// TIA Portal V20 program export: 0 tag tables, 0 data types, 52 data blocks, 105 code blocks (in call order from the OBs), 282 instance data blocks

DATA_BLOCK "Bypass"   // DB9
{ S7_Optimized_Access := 'TRUE' }
VERSION : 0.1
// stored: AutoNumber true, DBAccessibleFromOPCUA true, IsOnlyStoredInLoadMemory false, IsRetainMemResEnabled false, IsWriteProtectedInAS false, MemoryReserve 100
   VAR RETAIN
      Main_Panel { S7_SetPoint := 'True'} : "Safety_Bypass_MainPanel";
      Remote_Panel_1 : "Safety_Bypass_RemotePanel";
      Remote_Panel_2 { S7_SetPoint := 'True'} : "Safety_Bypass_RemotePanel";
      Remote_Panel_3 { S7_SetPoint := 'True'} : "Safety_Bypass_RemotePanel";
      Remote_Panel_4 { S7_SetPoint := 'True'} : "Safety_Bypass_RemotePanel";
      Remote_Panel_5 { S7_SetPoint := 'True'} : "Safety_Bypass_RemotePanel";
   END_VAR
BEGIN
   Main_Panel.Estop_Cabinet := FALSE;
END_DATA_BLOCK

DATA_BLOCK "Bypass_Safe"   // DB39, F_DB
{ S7_Optimized_Access := 'TRUE' }
VERSION : 0.1
// stored: AutoNumber true, DBAccessibleFromOPCUA true
   VAR
      Main_Panel : "F_Bypass_MainPanel";
      Remote_Panel_1 : "F_Bypass_RemotePanel";
      Remote_Panel_2 : "F_Bypass_RemotePanel";
      Remote_Panel_3 : "F_Bypass_RemotePanel";
      Remote_Panel_4 : "F_Bypass_RemotePanel";
      Remote_Panel_5 : "F_Bypass_RemotePanel";
   END_VAR
BEGIN
END_DATA_BLOCK

DATA_BLOCK "CNV_HMI"   // DB40
{ S7_Optimized_Access := 'TRUE' }
VERSION : 0.1
// stored: AutoNumber true, DBAccessibleFromOPCUA true, IsOnlyStoredInLoadMemory false, IsRetainMemResEnabled false, IsWriteProtectedInAS false, MemoryReserve 100
   VAR
      "Manual_Sfty_Stopper_Up(1)" : Array[1..5] of Bool;
      "Manual_Sfty_Stopper_Down(1)" : Array[1..5] of Bool;
      In_Out : Array[1..5] of Bool;
      ID : Array[1..5] of DInt;
      "Task_ID(1)" : Array[1..5] of UInt;
      Manual_Bwd : Array[1..5] of Bool;
      "Reset(1)" : Array[1..5] of Bool;
      "Pallet_Type(1)" : Array[1..5] of UInt;
      Manual_Fwd : Array[1..5] of Bool;
      Enable : Array[1..5] of Bool;
      "Pallet_Align_Right(1)" : Array[1..5] of Bool;
      "Enable(1)" : Array[1..5] of Bool;
      Pallet_Type : Array[1..5] of UInt;
      Pallet_Allignment : Array[1..5] of Bool;
      "Transfer_To_ID(1)" : Array[1..5] of DInt;
      Pallet_Align_Right : Array[1..5] of Bool;
      "Manual_Bwd(1)" : Array[1..5] of Bool;
      "Pallet_Align_Left(1)" : Array[1..5] of Bool;
      Reset : Array[1..5] of Bool;
      Stop : Array[1..5] of Bool;
      Pallet_Align_Center : Array[1..5] of Bool;
      "Stop(1)" : Array[1..5] of Bool;
      "Start_Transfer(1)" : Array[1..5] of Bool;
      Pallet_Align_Left : Array[1..5] of Bool;
      Start_Transfer : Array[1..5] of Bool;
      "ID(1)" : Array[1..5] of DInt;
      "Transfer_From_ID(1)" : Array[1..5] of DInt;
      "Manual_Fwd(1)" : Array[1..5] of Bool;
      Mode_Change : Array[1..5] of UInt;
      Transfer_To_ID : Array[1..5] of DInt;
      "Mode_Change(1)" : Array[1..5] of UInt;
      Transfer_From_ID : Array[1..5] of DInt;
      UpDown : Array[1..5] of UInt;
      Same_Cnv : Array[1..5] of Bool;
      CNV2_Selected : Array[1..5] of UInt;
      "Pallet_Allignment(1)" : Array[1..5] of Bool;
      "Occupied(1)" : Array[1..5] of Bool;
      Mode : Array[1..5] of UInt;
      "Running(1)" : Array[1..5] of Bool;
      "Enabled(1)" : Array[1..5] of Bool;
      Motor_Speed_Actual : Array[1..5] of UInt;
      Running : Array[1..5] of Bool;
      "SM_State(1)" : Array[1..5] of UInt;
      "Warning(1)" : Array[1..5] of UInt;
      Stopped : Array[1..5] of Bool;
      Enabled : Array[1..5] of Bool;
      Error : Array[1..5] of Bool;
      "Motor_Speed_Requested(1)" : Array[1..5] of UInt;
      Current_Task_ID : Array[1..5] of UInt;
      "Mode(1)" : Array[1..5] of UInt;
      "Current_Task_Type(1)" : Array[1..5] of UInt;
      Warning : Array[1..5] of UInt;
      "Current_Task_ID(1)" : Array[1..5] of UInt;
      Current_Task_Type : Array[1..5] of UInt;
      "Stopped(1)" : Array[1..5] of Bool;
      Motor_Direction : Array[1..5] of UInt;
      SM_State : Array[1..5] of UInt;
      "Ready_For_Task(1)" : Array[1..5] of Bool;
      Ready_For_Task : Array[1..5] of Bool;
      Occupied : Array[1..5] of Bool;
      "Error(1)" : Array[1..5] of Bool;
      Shuttle_in_place : Array[1..5] of Bool;
      Motor_Speed_Requested : Array[1..5] of UInt;
      "Motor_Direction(1)" : Array[1..5] of UInt;
      "Motor_Speed_Actual(1)" : Array[1..5] of UInt;
      "Shuttle_in_place(1)" : Array[1..5] of Bool;
      Motor_Ready : Array[1..5] of Bool;
      "Motor_Current_Actual(1)" : Array[1..5] of Real;
      Motor_Status : Array[1..5] of UInt;
      "Motor_Status(1)" : Array[1..5] of UInt;
      Motor_Current_Actual : Array[1..5] of Real;
      "Motor_Ready(1)" : Array[1..5] of Bool;
      Task_ID : Array[1..5] of UInt;
      Level_Selected : Array[1..5] of UInt;
      "UpDown(1)" : Array[1..5] of UInt;
      Motor_Actual_Torque : Array[1..5] of Real;
      "Motor_Actual_Torque(1)" : Array[1..5] of Real;
      Safety_OK : Array[1..5] of Bool;
      Reset_Comissioning : Array[1..5] of Bool;
      Charge_Commands : Array[1..5] of Bool;
      Charge_Cnv : Array[1..5] of Bool;
      Reset_All : Array[1..5] of Bool;
      Sdetect1 : Array[1..5] of Bool;
      Sdetect2 : Array[1..5] of Bool;
      "Sdetect1(1)" : Array[1..5] of Bool;
      "Sdetect2(1)" : Array[1..5] of Bool;
      "Rpd2(1)" : Array[1..5] of Bool;
      Center : Array[1..5] of Bool;
      "Rpd1(1)" : Array[1..5] of Bool;
      "Lpd2(1)" : Array[1..5] of Bool;
      "Lpd1(1)" : Array[1..5] of Bool;
      Rpd1 : Array[1..5] of Bool;
      Lpd1 : Array[1..5] of Bool;
      Rpd2 : Array[1..5] of Bool;
      "Right(1)" : Array[1..5] of Bool;
      Right : Array[1..5] of Bool;
      Left : Array[1..5] of Bool;
      "Left(1)" : Array[1..5] of Bool;
   END_VAR
BEGIN
END_DATA_BLOCK

DATA_BLOCK "Control_DB"   // DB69
{ S7_Optimized_Access := 'TRUE' }
VERSION : 0.1
// stored: AutoNumber true, DBAccessibleFromOPCUA true, IsOnlyStoredInLoadMemory false, IsRetainMemResEnabled false, IsWriteProtectedInAS false, MemoryReserve 100
   VAR
      ECnv_Sys { S7_SetPoint := 'True'} : Array[1..5] of "ECnv_Control";
      LCnv_Sys { S7_SetPoint := 'True'} : Array[1..5] of "Cnv_VTD_Control";
      VTD_Sys { S7_SetPoint := 'True'} : Array[1..5] of "VTD_Control";
      WCS_OPC_Control { S7_SetPoint := 'True'} : Array[1..5] of "WMS_OPC_UA";
      Shuttles_Position : Array[1..23] of Struct
         x : DInt;
         y : DInt;
         Charging : Bool;
      END_STRUCT;
      VTDBarcode_Station : Array[1..5] of "Barcode_Station_UDT";
      Pallet_ID_Received : Array[1..3] of Bool;
      Gate_Station : Array[1..12] of "Gate_Station_UDT";
   END_VAR
BEGIN
   LCnv_Sys[4].Cnv_Level[1..8].Cnv2.Safety_Stop_Cnrl.Inputs.DP_Extended := TRUE;
   LCnv_Sys[5].Cnv_Level[1..8].Cnv2.Safety_Stop_Cnrl.Inputs.DP_Extended := TRUE;
END_DATA_BLOCK

DATA_BLOCK "DB_Receive_Data_From_Logistex"   // DB900
{ S7_Optimized_Access := 'TRUE' }
VERSION : 0.1
// stored: AutoNumber false, DBAccessibleFromOPCUA true, IsOnlyStoredInLoadMemory false, IsRetainMemResEnabled false, IsWriteProtectedInAS false, MemoryReserve 100
   VAR
      J1310_Conv_Infeed : "Conv_Infeed";
      J1320_Conv_Infeed { S7_SetPoint := 'True'} : "Conv_Infeed";
      J1330_Conv_Infeed { S7_SetPoint := 'True'} : "Conv_Infeed";
      J1310_Conv_Oufeed { S7_SetPoint := 'True'} : "Conv_Outfeed";
      J1320_Conv_Oufeed { S7_SetPoint := 'True'} : "Conv_Outfeed";
      J1330_Conv_Oufeed { S7_SetPoint := 'True'} : "Conv_Outfeed";
      CNV_STATUS : Array[1..10] of Byte;
      PLC_STATUS : Struct
         Hardbit : Bool;
         "PLC_E-Stop" : Bool;
      END_STRUCT;
   END_VAR
BEGIN
END_DATA_BLOCK

DATA_BLOCK "DB_Send_Data_To_Logistex"   // DB901
{ S7_Optimized_Access := 'TRUE' }
VERSION : 0.1
// stored: AutoNumber false, DBAccessibleFromOPCUA true, IsOnlyStoredInLoadMemory false, IsRetainMemResEnabled false, IsWriteProtectedInAS false, MemoryReserve 100
   VAR
      VTD_J1310_INFEED : "VTD_Infeed";
      VTD_J1320_INFEED { S7_SetPoint := 'True'} : "VTD_Infeed";
      VTD_J1330_INFEED { S7_SetPoint := 'True'} : "VTD_Infeed";
      VTD_J1310_OUTFEED { S7_SetPoint := 'True'} : "VTD_Outfeed";
      VTD_J1320_OUTFEED { S7_SetPoint := 'True'} : "VTD_Outfeed";
      VTD_J1330_OUTFEED { S7_SetPoint := 'True'} : "VTD_Outfeed";
      VTD_STATUS : Array[1..10] of Byte;
      PLC_STATUS : Struct
         Hardbit : Bool;
         "PLC_E-Stop" : Bool;
      END_STRUCT;
      CONV_SPEED : Struct
         VTD_J1310_INF_SP : Int;
         VTD_J1310_OUF_SP : Int;
         VTD_J1320_INF_SP : Int;
         VTD_J1320_OUF_SP : Int;
         VTD_J1330_INF_SP_1 : Int;
         VTD_J1330_OUF_SP : Int;
      END_STRUCT;
   END_VAR
BEGIN
END_DATA_BLOCK

DATA_BLOCK "Force"   // DB12
{ S7_Optimized_Access := 'TRUE' }
VERSION : 0.1
// stored: AutoNumber true, DBAccessibleFromOPCUA true, IsOnlyStoredInLoadMemory false, IsRetainMemResEnabled false, IsWriteProtectedInAS false, MemoryReserve 100
   VAR
      "MAIN PANEL STACK LIGHT RED" : Bool;
      "MAIN PANEL STACK LIGHT AMBER" : Bool;
      "MAIN PANEL STACK LIGHT GREEN" : Bool;
      Remote_Panel : Array[1..5] of Struct
         "CX101_SFTY STOPPER ROTATE" : Bool;
         "CX102_SFTY STOPPER ROTATE" : Bool;
         "CX103_SFTY STOPPER ROTATE" : Bool;
         "CX104_SFTY STOPPER ROTATE" : Bool;
         "CX105_SFTY STOPPER ROTATE" : Bool;
         "CX106_SFTY STOPPER ROTATE" : Bool;
         "CX107_SFTY STOPPER ROTATE" : Bool;
         "CX108_SFTY STOPPER ROTATE" : Bool;
         "CX201_SFTY STOPPER ROTATE" : Bool;
         "CX202_SFTY STOPPER ROTATE" : Bool;
         "CX203_SFTY STOPPER ROTATE" : Bool;
         "CX204_SFTY STOPPER ROTATE" : Bool;
         "CX205_SFTY STOPPER ROTATE" : Bool;
         "CX206_SFTY STOPPER ROTATE" : Bool;
         "CX207_SFTY STOPPER ROTATE" : Bool;
         "CX208_SFTY STOPPER ROTATE" : Bool;
         "VTDx DOCKING PINS 1 RETRACT" : Bool;
         "VTDx DOCKING PINS 1 EXTEND" : Bool;
         "VTDx DOCKING PINS 2 EXTEND" : Bool;
         "VTDx DOCKING PINS 2 RETRACT" : Bool;
         "SCA X00Y STACK LIGHTS AMBER" : Bool;
         "SCA X00Y STACK LIGHTS GREEN" : Bool;
         "SCA X00Y STACK LIGHTS RED" : Bool;
         "EMERGENCY STOP RESET STATUS - ON(X)" : Bool;
      END_STRUCT;
   END_VAR
BEGIN
END_DATA_BLOCK

DATA_BLOCK "HMI_DB"   // DB21
{ S7_Optimized_Access := 'TRUE' }
VERSION : 0.1
// stored: AutoNumber true, DBAccessibleFromOPCUA true, IsOnlyStoredInLoadMemory false, IsRetainMemResEnabled false, IsWriteProtectedInAS false, MemoryReserve 100
   VAR
      Username : String := 'admin';
      Password : String := '12345';
      ScreenNo : Array[1..5] of UInt;
      ScreenNo_Main : UInt;
      System_Selected : Array[1..5] of UInt;
      Rem_Loc_Keys { ExternalAccessible := 'False'; ExternalVisible := 'False'; ExternalWritable := 'False'} : Array[1..5] of "Level_Keys_UDT";
   END_VAR
BEGIN
END_DATA_BLOCK

DATA_BLOCK "HMI_OrderTable"   // DB110
{ S7_Optimized_Access := 'TRUE' }
VERSION : 0.1
// stored: AutoNumber true, DBAccessibleFromOPCUA true, IsOnlyStoredInLoadMemory false, IsRetainMemResEnabled false, IsWriteProtectedInAS false, MemoryReserve 100
   VAR
      OrderTable : Array[0..9] of "OrderTable_UDT";
      State { S7_SetPoint := 'True'} : Array[0..9] of USInt;
      Index : Array[0..9] of Int;
      ScrollUp_PB : Bool;
      ScrollDown_PB : Bool;
      PlaceOrder_PB : Bool;
      PauseOrders_PB : Bool;
      ResumeOrder_PB : Bool;
      CancelOrder_PB : Bool;
      CancelThisOrder_PB : Bool;
      StartRow : Int;
      Device : USInt;
      PlacingNewOrder : Bool;
      PopUp_ErrorWindow_Active : Bool;
      PopUp_ErrorID : UInt;
      PopUp_Index : Int;
   END_VAR
BEGIN
END_DATA_BLOCK

DATA_BLOCK "HMI_OrderTable_1"   // DB137
{ S7_Optimized_Access := 'TRUE' }
VERSION : 0.1
// stored: AutoNumber true, DBAccessibleFromOPCUA true, IsOnlyStoredInLoadMemory false, IsRetainMemResEnabled false, IsWriteProtectedInAS false, MemoryReserve 100
   VAR
      OrderTable : Array[0..9] of "OrderTable_UDT";
      State { S7_SetPoint := 'True'} : Array[0..9] of USInt;
      Index : Array[0..9] of Int;
      ScrollUp_PB : Bool;
      ScrollDown_PB : Bool;
      PlaceOrder_PB : Bool;
      PauseOrders_PB : Bool;
      ResumeOrder_PB : Bool;
      CancelOrder_PB : Bool;
      CancelThisOrder_PB : Bool;
      StartRow : Int;
      Device : USInt;
      PlacingNewOrder : Bool;
      PopUp_ErrorWindow_Active : Bool;
      PopUp_ErrorID : UInt;
      PopUp_Index : Int;
   END_VAR
BEGIN
END_DATA_BLOCK

DATA_BLOCK "OrderTable_HMI"   // DB96
{ S7_Optimized_Access := 'TRUE' }
VERSION : 0.1
// stored: AutoNumber true, DBAccessibleFromOPCUA true, IsOnlyStoredInLoadMemory false, IsRetainMemResEnabled false, IsWriteProtectedInAS false, MemoryReserve 100
   VAR
      Start : Bool;
      Pause : Bool;
      Resume : Bool;
      Stop : Bool;
      "Manual order" : Bool;
      Transfer_From_To : Byte;
      "Send VTD Order" : Bool;
      "Send CNV Order" : Bool;
      "Pallet Type" : Byte;
      "Tower 1 Pallet Alignment" : Byte;
      "Tower 2 Pallet Alignment" : Byte;
      "Extractor Pallet Alignment" : Byte;
      "From level" : Byte;
      "To level" : Byte;
      "Testing Time" : UInt;
      "Numer of cycles" : Byte;
      Tower : Byte;
      Level : Byte;
      "Time Running" : UInt;
      Actual_Cycle : Byte;
      "Start Test Visibility" : Bool;
      "Stop Test Visibility" : Bool;
      "Pause Test Visibility" : Bool;
      "Resume Visibility" : Bool;
      "Clear Table Visibility" : Bool;
      "Pallet Type Visibility" : Bool;
      "Tower 1 Visibility" : Bool;
      "Tower 2 Visibility" : Bool;
      "Extractor Visibility" : Bool;
      Auto_Settings_Visibility : Bool;
      "ToExtractor Visibility" : Bool;
      "Manual order Visibility" : Bool;
      "Tower Visibility" : Bool;
      "Level Visibility" : Bool;
      "Send VTD Order Visibility" : Bool;
      "Send CNV Order Visibility" : Bool;
   END_VAR
BEGIN
END_DATA_BLOCK

DATA_BLOCK "OrderTable_HMI_1"   // DB99
{ S7_Optimized_Access := 'TRUE' }
VERSION : 0.1
// stored: AutoNumber true, DBAccessibleFromOPCUA true, IsOnlyStoredInLoadMemory false, IsRetainMemResEnabled false, IsWriteProtectedInAS false, MemoryReserve 100
   VAR
      Start : Bool;
      Pause : Bool;
      Resume : Bool;
      Stop : Bool;
      "Manual order" : Bool;
      Transfer_From_To : Byte;
      "Send VTD Order" : Bool;
      "Send CNV Order" : Bool;
      "Pallet Type" : Byte;
      "Tower 1 Pallet Alignment" : Byte;
      "Tower 2 Pallet Alignment" : Byte;
      "Extractor Pallet Alignment" : Byte;
      "From level" : Byte;
      "To level" : Byte;
      "Testing Time" : UInt;
      "Numer of cycles" : Byte;
      Tower : Byte;
      Level : Byte;
      "Time Running" : UInt;
      Actual_Cycle : Byte;
      "Start Test Visibility" : Bool;
      "Stop Test Visibility" : Bool;
      "Pause Test Visibility" : Bool;
      "Resume Visibility" : Bool;
      "Clear Table Visibility" : Bool;
      "Pallet Type Visibility" : Bool;
      "Tower 1 Visibility" : Bool;
      "Tower 2 Visibility" : Bool;
      "Extractor Visibility" : Bool;
      Auto_Settings_Visibility : Bool;
      "ToExtractor Visibility" : Bool;
      "Manual order Visibility" : Bool;
      "Tower Visibility" : Bool;
      "Level Visibility" : Bool;
      "Send VTD Order Visibility" : Bool;
      "Send CNV Order Visibility" : Bool;
      Clear_OT : Bool;
   END_VAR
BEGIN
END_DATA_BLOCK

DATA_BLOCK "Overhang_IO_DB"   // DB439, F_DB
{ S7_Optimized_Access := 'TRUE' }
VERSION : 0.1
// stored: AutoNumber true, DBAccessibleFromOPCUA true
   VAR
      ECnv_1 : "F_ECnv_Overhang";
      ECnv_2 : "F_ECnv_Overhang";
      ECnv_3 : "F_ECnv_Overhang";
      ECnv_4 : "F_ECnv_Overhang";
      ECnv_5 : "F_ECnv_Overhang";
   END_VAR
BEGIN
END_DATA_BLOCK

DATA_BLOCK "PopUp_Screens_1"   // DB51
{ S7_Optimized_Access := 'TRUE' }
VERSION : 0.1
// stored: AutoNumber true, DBAccessibleFromOPCUA true, IsOnlyStoredInLoadMemory false, IsRetainMemResEnabled false, IsWriteProtectedInAS false, MemoryReserve 100
   VAR
      LE_Speed : Array[1..6] of DInt;
      LE_Warnings : Array[1..6] of Byte;
      LE_Status : Array[1..6] of Bool;
      LE_Quality_Value : Array[1..6] of Int;
      LE_X_Unsafe_Position : Array[1..6] of UInt;
      LE_Quality_Decoded_Codes : Array[1..6] of UInt;
      LE_Bypass : Array[1..6] of DInt;
      AE_Speed : Array[1..6] of DInt;
      AE_Status_2 : Array[1..6] of UInt;
      AE_Control_Word_2 : Array[1..6] of UInt;
      AE_Position_1 : Array[1..6] of Bool;
      AE_Position_2 : Array[1..6] of Bool;
      AE_Status_1 : Array[1..6] of Bool;
      AE_Control_Word_1 : Array[1..6] of Bool;
      BCD_Disable_Trigger_HMI : Array[1..6] of Bool;
      BCD_Enable_Trigger_HMI : Array[1..6] of Bool;
      BCD_Error_HMI : Array[1..6] of Bool;
      BCD_Start_Comm_Test_HMI : Array[1..6] of Bool;
      BCD_Test_Ok_HMI : Array[1..6] of Bool;
      BCD_Execute_Function : Array[1..6] of Bool;
      BCD_RdDone : Array[1..6] of Bool;
      BCD_ReqDone : Array[1..6] of Bool;
      BCD_ReqBusy : Array[1..6] of Bool;
   END_VAR
BEGIN
END_DATA_BLOCK

DATA_BLOCK "PopUps_DB"   // DB38
{ S7_Optimized_Access := 'TRUE' }
VERSION : 0.1
// stored: AutoNumber false, DBAccessibleFromOPCUA true, IsOnlyStoredInLoadMemory false, IsRetainMemResEnabled false, IsWriteProtectedInAS false, MemoryReserve 100
   VAR
      Buffer_Cnv_Settings_1 : "Buffer_Cnv_Settings";
      Buffer_Cnv_Settings_2 { S7_SetPoint := 'True'} : "Buffer_Cnv_Settings";
      ECnv_Settings { S7_SetPoint := 'True'} : "ECnv_Settings";
      VTD_Settings { S7_SetPoint := 'True'} : "VTD_Settings";
      Shuttle_MQTT_Settings { S7_SetPoint := 'True'} : "MQTT_Settings";
      Sick_Lector_Reseult : String;
   END_VAR
BEGIN
END_DATA_BLOCK

DATA_BLOCK "PopUps_DB_1"   // DB20
{ S7_Optimized_Access := 'TRUE' }
VERSION : 0.1
// stored: AutoNumber true, DBAccessibleFromOPCUA true, IsOnlyStoredInLoadMemory false, IsRetainMemResEnabled false, IsWriteProtectedInAS false, MemoryReserve 100
   VAR
      Buffer_Cnv_Settings_1 : Array[1..5] of "Buffer_Cnv_Settings";
      Buffer_Cnv_Settings_2 { S7_SetPoint := 'True'} : Array[1..5] of "Buffer_Cnv_Settings";
      ECnv_Settings { S7_SetPoint := 'True'} : Array[1..5] of "ECnv_Settings";
      VTD_Settings { S7_SetPoint := 'True'} : Array[1..5] of "VTD_Settings";
      Shuttle_MQTT_Settings { S7_SetPoint := 'True'} : "MQTT_Settings";
      Sick_Lector_Reseult : Array[1..5] of String;
      Save_Settings { S7_SetPoint := 'True'} : Array[1..5] of Bool;
      Absolute_Encoder : Array[1..5] of Struct
         AE_Control_Word_1 : UInt;
         AE_Control_Word_2 : UInt;
         AE_Status_1 : UInt;
         AE_Status_2 : UInt;
         AE_Position_1 : DInt;
         AE_Position_2 : DInt;
         AE_Speed : Int;
      END_STRUCT;
      Lector_Barcode : Array[1..5] of Struct
         BCD_Test_Comm : Bool;
         BCD_Disable_Trigger : Bool;
         BCD_Enable_Trigger : Bool;
         BCD_Execute_Function : Bool;
         BCD_Test_Ok : Bool;
         BCD_Error : Bool;
         BCD_RdDone : Bool;
         BCD_ReqDone : Bool;
         BCD_ReqBusy : Bool;
         Lector_Reseult : String;
      END_STRUCT;
      Linear_Encoder : Array[1..5] of Struct
         LE_X_Unsafe_Position : DInt;
         LE_Speed : Int;
         LE_Warnings : Int;
         LE_Bypass : Bool;
         LE_Status : UInt;
      END_STRUCT;
      Trend : Array[1..5] of Struct
         Motor_SetPoint : UInt;
         Motor_Actual_Current : Real;
         Motor_Actual_Speed : UInt;
      END_STRUCT;
   END_VAR
BEGIN
   Shuttle_MQTT_Settings.MQTT_Con_Params.hwId := 64;
   Shuttle_MQTT_Settings.MQTT_Con_Params.broker := '10.0.34.2';
   Shuttle_MQTT_Settings.Client_ID := WSTRING#'PLC';
   Shuttle_MQTT_Settings.Username := WSTRING#'Devin';
   Shuttle_MQTT_Settings.Password := WSTRING#'1';
   Shuttle_MQTT_Settings.Retain := TRUE;
END_DATA_BLOCK

DATA_BLOCK "SICK_AFx60_Data_DB"   // DB120
{ S7_Optimized_Access := 'TRUE' }
VERSION : 0.1
// stored: AutoNumber true, DBAccessibleFromOPCUA true, IsOnlyStoredInLoadMemory false, IsRetainMemResEnabled false, IsWriteProtectedInAS false, MemoryReserve 100
   VAR
      "Absolute Encoder 1" { S7_SetPoint := 'True'} : "ST_SICK_AFx60";
      "Absolute Encoder 2" { S7_SetPoint := 'True'} : "ST_SICK_AFx60";
      "Absolute Encoder 3" { S7_SetPoint := 'True'} : "ST_SICK_AFx60";
      "Absolute Encoder 4" { S7_SetPoint := 'True'} : "ST_SICK_AFx60";
      "Absolute Encoder 5" { S7_SetPoint := 'True'} : "ST_SICK_AFx60";
   END_VAR
BEGIN
END_DATA_BLOCK

DATA_BLOCK "SICK_Lector_DB_1"   // DB46
{ S7_Optimized_Access := 'TRUE' }
VERSION : 0.1
// stored: AutoNumber true, DBAccessibleFromOPCUA true, IsOnlyStoredInLoadMemory false, IsRetainMemResEnabled false, IsWriteProtectedInAS false, MemoryReserve 100
   VAR
      Barcode_Result : String;
      Test_OK : Bool;
      HWInputIdent : HW_IO := 554;
      HWInputLength : USInt := 32;
      HWOutputIdent : HW_IO := 555;
      HWOutputLength : USInt := 32;
      CANId : USInt := 0;
      TOut : Time := T#10S;
      Req : Bool := FALSE;
      TriggerOn : Bool := FALSE;
      TriggerOff : Bool := FALSE;
      Matchcode : Bool := FALSE;
      SavePermanent : Bool := FALSE;
      ComTest : Bool := FALSE;
      FreeCommand : Bool := FALSE;
      Data : "ST_SICK_Lector_CLV6xx";
      RdDone { S7_SetPoint := 'True'} : Bool := FALSE;
      ReqDone : Bool := FALSE;
      ReqBusy : Bool := FALSE;
      Error : Bool := TRUE;
      Errorcode : DWord := 16#0000_0015;
   END_VAR
BEGIN
   Data.Matchcode.sName := '';
   Data.Matchcode.nCodeType := ' ';
   Data.Matchcode.iMinMaxLength := 0;
   Data.Matchcode.sContent := '';
   Data.FreeCommand.sCommand := '';
   Data.FreeCommand.sResult := '';
   Data.ReadingResult.iCounter := 0;
   Data.ReadingResult.iLength := 0;
   Data.ReadingResult.arrResult[1..200] := 16#00;
END_DATA_BLOCK

DATA_BLOCK "SICK_Lector_DB_2"   // DB309
{ S7_Optimized_Access := 'TRUE' }
VERSION : 0.1
// stored: AutoNumber true, DBAccessibleFromOPCUA true, IsOnlyStoredInLoadMemory false, IsRetainMemResEnabled false, IsWriteProtectedInAS false, MemoryReserve 100
   VAR
      Barcode_Result : String;
      Test_OK : Bool;
      HWInputIdent : HW_IO := 554;
      HWInputLength : USInt := 32;
      HWOutputIdent : HW_IO := 555;
      HWOutputLength : USInt := 32;
      CANId : USInt := 0;
      TOut : Time := T#10S;
      Req : Bool := FALSE;
      TriggerOn : Bool := FALSE;
      TriggerOff : Bool := FALSE;
      Matchcode : Bool := FALSE;
      SavePermanent : Bool := FALSE;
      ComTest : Bool := FALSE;
      FreeCommand : Bool := FALSE;
      Data : "ST_SICK_Lector_CLV6xx";
      RdDone { S7_SetPoint := 'True'} : Bool := FALSE;
      ReqDone : Bool := FALSE;
      ReqBusy : Bool := FALSE;
      Error : Bool := TRUE;
      Errorcode : DWord := 16#0000_0015;
   END_VAR
BEGIN
   Data.Matchcode.sName := '';
   Data.Matchcode.nCodeType := ' ';
   Data.Matchcode.iMinMaxLength := 0;
   Data.Matchcode.sContent := '';
   Data.FreeCommand.sCommand := '';
   Data.FreeCommand.sResult := '';
   Data.ReadingResult.iCounter := 0;
   Data.ReadingResult.iLength := 0;
   Data.ReadingResult.arrResult[1..200] := 16#00;
END_DATA_BLOCK

DATA_BLOCK "SICK_Lector_DB_3"   // DB310
{ S7_Optimized_Access := 'TRUE' }
VERSION : 0.1
// stored: AutoNumber true, DBAccessibleFromOPCUA true, IsOnlyStoredInLoadMemory false, IsRetainMemResEnabled false, IsWriteProtectedInAS false, MemoryReserve 100
   VAR
      Barcode_Result : String;
      Test_OK : Bool;
      HWInputIdent : HW_IO := 554;
      HWInputLength : USInt := 32;
      HWOutputIdent : HW_IO := 555;
      HWOutputLength : USInt := 32;
      CANId : USInt := 0;
      TOut : Time := T#10S;
      Req : Bool := FALSE;
      TriggerOn : Bool := FALSE;
      TriggerOff : Bool := FALSE;
      Matchcode : Bool := FALSE;
      SavePermanent : Bool := FALSE;
      ComTest : Bool := FALSE;
      FreeCommand : Bool := FALSE;
      Data : "ST_SICK_Lector_CLV6xx";
      RdDone { S7_SetPoint := 'True'} : Bool := FALSE;
      ReqDone : Bool := FALSE;
      ReqBusy : Bool := FALSE;
      Error : Bool := TRUE;
      Errorcode : DWord := 16#0000_0015;
   END_VAR
BEGIN
   Data.Matchcode.sName := '';
   Data.Matchcode.nCodeType := ' ';
   Data.Matchcode.iMinMaxLength := 0;
   Data.Matchcode.sContent := '';
   Data.FreeCommand.sCommand := '';
   Data.FreeCommand.sResult := '';
   Data.ReadingResult.iCounter := 0;
   Data.ReadingResult.iLength := 0;
   Data.ReadingResult.arrResult[1..200] := 16#00;
END_DATA_BLOCK

DATA_BLOCK "SICK_Lector_DB_4"   // DB307
{ S7_Optimized_Access := 'TRUE' }
VERSION : 0.1
// stored: AutoNumber true, DBAccessibleFromOPCUA true, IsOnlyStoredInLoadMemory false, IsRetainMemResEnabled false, IsWriteProtectedInAS false, MemoryReserve 100
   VAR
      Barcode_Result : String;
      Test_OK : Bool;
      HWInputIdent : HW_IO := 554;
      HWInputLength : USInt := 32;
      HWOutputIdent : HW_IO := 555;
      HWOutputLength : USInt := 32;
      CANId : USInt := 0;
      TOut : Time := T#10S;
      Req : Bool := FALSE;
      TriggerOn : Bool := FALSE;
      TriggerOff : Bool := FALSE;
      Matchcode : Bool := FALSE;
      SavePermanent : Bool := FALSE;
      ComTest : Bool := FALSE;
      FreeCommand : Bool := FALSE;
      Data : "ST_SICK_Lector_CLV6xx";
      RdDone { S7_SetPoint := 'True'} : Bool := FALSE;
      ReqDone : Bool := FALSE;
      ReqBusy : Bool := FALSE;
      Error : Bool := TRUE;
      Errorcode : DWord := 16#0000_0015;
   END_VAR
BEGIN
   Data.Matchcode.sName := '';
   Data.Matchcode.nCodeType := ' ';
   Data.Matchcode.iMinMaxLength := 0;
   Data.Matchcode.sContent := '';
   Data.FreeCommand.sCommand := '';
   Data.FreeCommand.sResult := '';
   Data.ReadingResult.iCounter := 0;
   Data.ReadingResult.iLength := 0;
   Data.ReadingResult.arrResult[1..200] := 16#00;
END_DATA_BLOCK

DATA_BLOCK "SICK_Lector_DB_5"   // DB308
{ S7_Optimized_Access := 'TRUE' }
VERSION : 0.1
// stored: AutoNumber true, DBAccessibleFromOPCUA true, IsOnlyStoredInLoadMemory false, IsRetainMemResEnabled false, IsWriteProtectedInAS false, MemoryReserve 100
   VAR
      Barcode_Result : String;
      Test_OK : Bool;
      HWInputIdent : HW_IO := 554;
      HWInputLength : USInt := 32;
      HWOutputIdent : HW_IO := 555;
      HWOutputLength : USInt := 32;
      CANId : USInt := 0;
      TOut : Time := T#10S;
      Req : Bool := FALSE;
      TriggerOn : Bool := FALSE;
      TriggerOff : Bool := FALSE;
      Matchcode : Bool := FALSE;
      SavePermanent : Bool := FALSE;
      ComTest : Bool := FALSE;
      FreeCommand : Bool := FALSE;
      Data : "ST_SICK_Lector_CLV6xx";
      RdDone { S7_SetPoint := 'True'} : Bool := FALSE;
      ReqDone : Bool := FALSE;
      ReqBusy : Bool := FALSE;
      Error : Bool := TRUE;
      Errorcode : DWord := 16#0000_0015;
   END_VAR
BEGIN
   Data.Matchcode.sName := '';
   Data.Matchcode.nCodeType := ' ';
   Data.Matchcode.iMinMaxLength := 0;
   Data.Matchcode.sContent := '';
   Data.FreeCommand.sCommand := '';
   Data.FreeCommand.sResult := '';
   Data.ReadingResult.iCounter := 0;
   Data.ReadingResult.iLength := 0;
   Data.ReadingResult.arrResult[1..200] := 16#00;
END_DATA_BLOCK

DATA_BLOCK "Safety_Communication"   // DB1000
{ S7_Optimized_Access := 'TRUE' }
VERSION : 0.1
// stored: AutoNumber false, DBAccessibleFromOPCUA true, IsOnlyStoredInLoadMemory false, IsRetainMemResEnabled false, IsWriteProtectedInAS false, MemoryReserve 100
   VAR
      RCV_ARRAY : Array[0..26] of Byte;
      ACK_SEND_ARRAY : Array[0..21] of Byte;
      SEND_ARRAY : Array[0..26] of Byte;
      ACK_RCV_ARRAY : Array[0..21] of Byte;
   END_VAR
BEGIN
END_DATA_BLOCK

DATA_BLOCK "Screen_DB"   // DB23
{ S7_Optimized_Access := 'TRUE' }
VERSION : 0.1
// stored: AutoNumber true, DBAccessibleFromOPCUA true, IsOnlyStoredInLoadMemory false, IsRetainMemResEnabled false, IsWriteProtectedInAS false, MemoryReserve 100
   VAR
      Settings_ActivePopUp : USInt;
      Alarms_ActiveTable : USInt;
      MainTemplate_ErrorActive : Bool;
      MainTemplate_ErrorCount : USInt;
      MainTemplate_Background : USInt;
      EmptyTemplate_Background : USInt;
      Charge_VTD : Bool;
      Charge_Cnv : Bool;
      Charge_VTD_Commands : Bool;
      Charge_Cnv_Commands : Bool;
      Charge_OT : Bool;
      Shuttle : "Shuttle_MQTT_Status_Msg";
      Shuttle_Select : USInt;
      VTD_Barcode : String;
      VTD_Barcode_Visu : Bool;
      OrderProcessing : Array[1..5] of String;
   END_VAR
BEGIN
END_DATA_BLOCK

DATA_BLOCK "Screen_DB_1"   // DB54
{ S7_Optimized_Access := 'TRUE' }
VERSION : 0.1
// stored: AutoNumber true, DBAccessibleFromOPCUA true, IsOnlyStoredInLoadMemory false, IsRetainMemResEnabled false, IsWriteProtectedInAS false, MemoryReserve 100
   VAR
      Charge_VTD_Commands : Array[1..5] of Bool;
      Shuttle : "Shuttle_MQTT_Status_Msg";
      Reset_All : Array[1..5] of Bool;
      Shuttle_Level_Selected : Array[1..5] of UInt;
      Charge_Shuttle_Commands : Array[1..5] of Bool;
      Shuttle_Select : Array[1..5] of USInt;
      Charge_OT { S7_SetPoint := 'True'} : Array[1..5] of Bool;
      OrderTable_Selected : Array[1..5] of UInt;
      Automatic_Button : Array[1..5] of Bool;
      All_In_Automatic : Array[1..5] of Bool;
      System_Error : Array[1..5] of Bool;
      Reset_Comissioning : Array[1..5] of Bool;
      Alarms_ActiveTable : Array[1..5] of USInt;
      Charger_1 : Array[1..5] of Bool;
      Charger_2 : Array[1..5] of Bool;
      Charger_3 : Array[1..5] of Bool;
      Shuttle_Charge_Buttons : Array[1..5] of Bool;
      Alarm_Current_Buttons : Array[1..5] of Bool;
      Alarm_History_Buttons : Array[1..5] of Bool;
      MainTemplate_Background : Array[1..5] of USInt;
      Settings_ActivePopUp : Array[1..5] of USInt;
      MainTemplate_ErrorActive : Array[1..5] of Bool;
      MainTemplate_ErrorCount : Array[1..5] of USInt;
      EmptyTemplate_Background : Array[1..5] of USInt;
      Charge_VTD : Array[1..5] of Bool;
      Charge_Cnv : Array[1..5] of Bool;
      Charge_Cnv_Commands : Array[1..5] of Bool;
   END_VAR
BEGIN
   Charger_1[1..5] := false;
END_DATA_BLOCK

DATA_BLOCK "Settings_DB"   // DB71
{ S7_Optimized_Access := 'TRUE' }
VERSION : 0.1
// stored: AutoNumber true, DBAccessibleFromOPCUA true, IsOnlyStoredInLoadMemory false, IsRetainMemResEnabled false, IsWriteProtectedInAS false, MemoryReserve 100
   VAR RETAIN
      VTD_Sys : Array[1..5] of "VTD_Settings";
      ECnv_Sys : Array[1..5] of "ECnv_Settings";
      LCnv_Sys : Array[1..5] of "Cnv_VTD_Settings";
      Shuttle_MQTT : "MQTT_Settings";
      System : "System_Settings";
   END_VAR
   VAR
      Chain_Slack_Time { S7_SetPoint := 'True'} : Time := t#200ms;
   END_VAR
BEGIN
   VTD_Sys[1].ID := 1;
   VTD_Sys[2].ID := 2;
   VTD_Sys[3].ID := 3;
   VTD_Sys[4].ID := 4;
   VTD_Sys[5].ID := 5;
   VTD_Sys[1..5].Lowest_Level := 1;
   VTD_Sys[1..5].Highest_Level := 8;
   VTD_Sys[1..3].VTD_Max_Heigh := 16500;
   VTD_Sys[4..5].VTD_Max_Heigh := 17000;
   VTD_Sys[1].VTD_Min_Height := 55;
   VTD_Sys[2].VTD_Min_Height := 0;
   VTD_Sys[3].VTD_Min_Height := 45;
   VTD_Sys[4..5].VTD_Min_Height := 0;
   VTD_Sys[1..5].VTD_Level_Granularity := 20;
   VTD_Sys[1..5].Dft_Level_Offset_LE := 0;
   VTD_Sys[1..5].Dft_Level_Offset_AE := 0;
   VTD_Sys[1..5].Teach_Speed := 0;
   VTD_Sys[1..5].Creep_Speed := 3;
   VTD_Sys[1].Slow_Speed := 5;
   VTD_Sys[2..5].Slow_Speed := 15;
   VTD_Sys[1..5].Slow_Calib_Speed := 10;
   VTD_Sys[1..5].Loaded_Speed := 50;
   VTD_Sys[1..5].Shuttle_Speed := 50;
   VTD_Sys[1..5].Pallet_Speed := 100;
   VTD_Sys[1..5].Empty_Speed := 100;
   VTD_Sys[1..5].Dock_speed := 5;
   VTD_Sys[1..5].Manual_Speed := 15;
   VTD_Sys[1..5].Slowdown_Count_LE := 700;
   VTD_Sys[1].Creep_Count_LE := 60;
   VTD_Sys[2].Creep_Count_LE := 50;
   VTD_Sys[3..5].Creep_Count_LE := 60;
   VTD_Sys[1..5].Slowdown_Count_AE := 700;
   VTD_Sys[1..5].Creep_Count_AE := 60;
   VTD_Sys[1..5].Encoder_Delta_W1 := 0.0;
   VTD_Sys[1..5].Encoder_Delta_W2 := 0.0;
   VTD_Sys[1..5].AE_Ratio := 0.0;
   VTD_Sys[1].Encoder_Delta_Warning := 80.0;
   VTD_Sys[2..5].Encoder_Delta_Warning := 50.0;
   VTD_Sys[1..5].Encoder_Delta_Error := 200.0;
   VTD_Sys[1..5].Transfer_Timeout_Up := 50;
   VTD_Sys[1..5].Transfer_Timeout_Down := 45;
   VTD_Sys[1..5].Lockpins_Timeout_Extend := 3000;
   VTD_Sys[1..5].Lockpins_Timeout_Retract := 3000;
   VTD_Sys[1].Level_Detect_Timeout := 500;
   VTD_Sys[2].Level_Detect_Timeout := 900;
   VTD_Sys[3..5].Level_Detect_Timeout := 500;
   VTD_Sys[1..5].Teach_Timeout := 600;
   VTD_Sys[1].Chain_Slack_Timeout := 750;
   VTD_Sys[2].Chain_Slack_Timeout := 500;
   VTD_Sys[3].Chain_Slack_Timeout := 600;
   VTD_Sys[4].Chain_Slack_Timeout := 500;
   VTD_Sys[5].Chain_Slack_Timeout := 1600;
   VTD_Sys[1].Level_Detect_LE := 3.0;
   VTD_Sys[2].Level_Detect_LE := 2.0;
   VTD_Sys[3..5].Level_Detect_LE := 3.0;
   VTD_Sys[1..5].Acc_Range_1 := 60;
   VTD_Sys[1..5].Acc_Range_2 := 70;
   VTD_Sys[1..5].Acc_Range_3 := 80;
   VTD_Sys[1..5].Weight_Range_1 := 250;
   VTD_Sys[1..5].Weight_Range_2 := 500;
   VTD_Sys[1..5].Weight_Range_3 := 750;
   VTD_Sys[1].G120_Hardware_ID := 475;
   VTD_Sys[2].G120_Hardware_ID := 959;
   VTD_Sys[3].G120_Hardware_ID := 1363;
   VTD_Sys[4].G120_Hardware_ID := 1767;
   VTD_Sys[5].G120_Hardware_ID := 2075;
   VTD_Sys[1].Teach_Values.Levels_LE[1] := 58.0;
   VTD_Sys[1].Teach_Values.Levels_LE[2] := 2525.0;
   VTD_Sys[1].Teach_Values.Levels_LE[3] := 4722.0;
   VTD_Sys[1].Teach_Values.Levels_LE[4] := 6927.0;
   VTD_Sys[1].Teach_Values.Levels_LE[5] := 9276.0;
   VTD_Sys[1].Teach_Values.Levels_LE[6] := 11627.0;
   VTD_Sys[1].Teach_Values.Levels_LE[7] := 13978.0;
   VTD_Sys[1].Teach_Values.Levels_LE[8] := 16325.0;
   VTD_Sys[2].Teach_Values.Levels_LE[1] := 63.0;
   VTD_Sys[2].Teach_Values.Levels_LE[2] := 2546.0;
   VTD_Sys[2].Teach_Values.Levels_LE[3] := 4744.0;
   VTD_Sys[2].Teach_Values.Levels_LE[4] := 6944.0;
   VTD_Sys[2].Teach_Values.Levels_LE[5] := 9291.0;
   VTD_Sys[2].Teach_Values.Levels_LE[6] := 11641.0;
   VTD_Sys[2].Teach_Values.Levels_LE[7] := 13993.0;
   VTD_Sys[2].Teach_Values.Levels_LE[8] := 16347.0;
   VTD_Sys[3].Teach_Values.Levels_LE[1] := 49.0;
   VTD_Sys[3].Teach_Values.Levels_LE[2] := 2524.0;
   VTD_Sys[3].Teach_Values.Levels_LE[3] := 4726.0;
   VTD_Sys[3].Teach_Values.Levels_LE[4] := 6923.0;
   VTD_Sys[3].Teach_Values.Levels_LE[5] := 9273.0;
   VTD_Sys[3].Teach_Values.Levels_LE[6] := 11623.0;
   VTD_Sys[3].Teach_Values.Levels_LE[7] := 13972.0;
   VTD_Sys[3].Teach_Values.Levels_LE[8] := 16328.0;
   VTD_Sys[4].Teach_Values.Levels_LE[1] := 161.0;
   VTD_Sys[4].Teach_Values.Levels_LE[2] := 2608.0;
   VTD_Sys[4].Teach_Values.Levels_LE[3] := 4807.0;
   VTD_Sys[4].Teach_Values.Levels_LE[4] := 7009.0;
   VTD_Sys[4].Teach_Values.Levels_LE[5] := 9358.0;
   VTD_Sys[4].Teach_Values.Levels_LE[6] := 11709.0;
   VTD_Sys[4].Teach_Values.Levels_LE[7] := 14057.0;
   VTD_Sys[4].Teach_Values.Levels_LE[8] := 16406.0;
   VTD_Sys[5].Teach_Values.Levels_LE[1] := 168.0;
   VTD_Sys[5].Teach_Values.Levels_LE[2] := 2609.0;
   VTD_Sys[5].Teach_Values.Levels_LE[3] := 4808.0;
   VTD_Sys[5].Teach_Values.Levels_LE[4] := 7007.0;
   VTD_Sys[5].Teach_Values.Levels_LE[5] := 9358.0;
   VTD_Sys[5].Teach_Values.Levels_LE[6] := 11705.0;
   VTD_Sys[5].Teach_Values.Levels_LE[7] := 14056.0;
   VTD_Sys[5].Teach_Values.Levels_LE[8] := 16404.0;
   VTD_Sys[1].Teach_Values.Levels_AE[1..8] := 0;
   VTD_Sys[2].Teach_Values.Levels_AE[1..8] := 0;
   VTD_Sys[3].Teach_Values.Levels_AE[1..8] := 0;
   VTD_Sys[4].Teach_Values.Levels_AE[1..8] := 0;
   VTD_Sys[5].Teach_Values.Levels_AE[1..8] := 0;
   ECnv_Sys[1].ID := 120101;
   ECnv_Sys[2].ID := 120102;
   ECnv_Sys[3].ID := 120203;
   ECnv_Sys[4].ID := 120104;
   ECnv_Sys[5].ID := 120105;
   ECnv_Sys[1].Barcode_ID := 1;
   ECnv_Sys[2].Barcode_ID := 2;
   ECnv_Sys[3].Barcode_ID := 3;
   ECnv_Sys[4].Barcode_ID := 4;
   ECnv_Sys[5].Barcode_ID := 5;
   ECnv_Sys[1..2].Cnv_Level := 1;
   ECnv_Sys[3].Cnv_Level := 2;
   ECnv_Sys[4..5].Cnv_Level := 1;
   ECnv_Sys[1..5].TC_Time := 20;
   ECnv_Sys[1..5].Transfer_Time := 20;
   ECnv_Sys[1..5].Pallet_Align_Time := 20;
   ECnv_Sys[1..5].Slow_Speed := 11;
   ECnv_Sys[1..5].Full_Speed := 100;
   ECnv_Sys[1..5].Manual_Speed := 40;
   ECnv_Sys[1..5].Timer_Check_Pallet_Time := 750;
   ECnv_Sys[1].G120_Hardware_ID := 488;
   ECnv_Sys[2].G120_Hardware_ID := 968;
   ECnv_Sys[3].G120_Hardware_ID := 1372;
   ECnv_Sys[4].G120_Hardware_ID := 1776;
   ECnv_Sys[5].G120_Hardware_ID := 2084;
   LCnv_Sys[1].Cnv_Level[1].Cnv1.ID := 100101;
   LCnv_Sys[1].Cnv_Level[2].Cnv1.ID := 100201;
   LCnv_Sys[1].Cnv_Level[3].Cnv1.ID := 100301;
   LCnv_Sys[1].Cnv_Level[4].Cnv1.ID := 100401;
   LCnv_Sys[1].Cnv_Level[5].Cnv1.ID := 100501;
   LCnv_Sys[1].Cnv_Level[6].Cnv1.ID := 100601;
   LCnv_Sys[1].Cnv_Level[7].Cnv1.ID := 100701;
   LCnv_Sys[1].Cnv_Level[8].Cnv1.ID := 100801;
   LCnv_Sys[2].Cnv_Level[1].Cnv1.ID := 100102;
   LCnv_Sys[2].Cnv_Level[2].Cnv1.ID := 100202;
   LCnv_Sys[2].Cnv_Level[3].Cnv1.ID := 100302;
   LCnv_Sys[2].Cnv_Level[4].Cnv1.ID := 100402;
   LCnv_Sys[2].Cnv_Level[5].Cnv1.ID := 100502;
   LCnv_Sys[2].Cnv_Level[6].Cnv1.ID := 100602;
   LCnv_Sys[2].Cnv_Level[7].Cnv1.ID := 100702;
   LCnv_Sys[2].Cnv_Level[8].Cnv1.ID := 100802;
   LCnv_Sys[3].Cnv_Level[1].Cnv1.ID := 100103;
   LCnv_Sys[3].Cnv_Level[2].Cnv1.ID := 100203;
   LCnv_Sys[3].Cnv_Level[3].Cnv1.ID := 100303;
   LCnv_Sys[3].Cnv_Level[4].Cnv1.ID := 100403;
   LCnv_Sys[3].Cnv_Level[5].Cnv1.ID := 100503;
   LCnv_Sys[3].Cnv_Level[6].Cnv1.ID := 100603;
   LCnv_Sys[3].Cnv_Level[7].Cnv1.ID := 100703;
   LCnv_Sys[3].Cnv_Level[8].Cnv1.ID := 100803;
   LCnv_Sys[4].Cnv_Level[1].Cnv1.ID := 100104;
   LCnv_Sys[4].Cnv_Level[2].Cnv1.ID := 100204;
   LCnv_Sys[4].Cnv_Level[3].Cnv1.ID := 100304;
   LCnv_Sys[4].Cnv_Level[4].Cnv1.ID := 100404;
   LCnv_Sys[4].Cnv_Level[5].Cnv1.ID := 100504;
   LCnv_Sys[4].Cnv_Level[6].Cnv1.ID := 100604;
   LCnv_Sys[4].Cnv_Level[7].Cnv1.ID := 100704;
   LCnv_Sys[4].Cnv_Level[8].Cnv1.ID := 100804;
   LCnv_Sys[5].Cnv_Level[1].Cnv1.ID := 100105;
   LCnv_Sys[5].Cnv_Level[2].Cnv1.ID := 100205;
   LCnv_Sys[5].Cnv_Level[3].Cnv1.ID := 100305;
   LCnv_Sys[5].Cnv_Level[4].Cnv1.ID := 100405;
   LCnv_Sys[5].Cnv_Level[5].Cnv1.ID := 100505;
   LCnv_Sys[5].Cnv_Level[6].Cnv1.ID := 100605;
   LCnv_Sys[5].Cnv_Level[7].Cnv1.ID := 100705;
   LCnv_Sys[5].Cnv_Level[8].Cnv1.ID := 100805;
   LCnv_Sys[1].Cnv_Level[1].Cnv1.Barcode_ID := 6;
   LCnv_Sys[1].Cnv_Level[2].Cnv1.Barcode_ID := 14;
   LCnv_Sys[1].Cnv_Level[3].Cnv1.Barcode_ID := 22;
   LCnv_Sys[1].Cnv_Level[4].Cnv1.Barcode_ID := 30;
   LCnv_Sys[1].Cnv_Level[5].Cnv1.Barcode_ID := 38;
   LCnv_Sys[1].Cnv_Level[6].Cnv1.Barcode_ID := 46;
   LCnv_Sys[1].Cnv_Level[7].Cnv1.Barcode_ID := 54;
   LCnv_Sys[1].Cnv_Level[8].Cnv1.Barcode_ID := 62;
   LCnv_Sys[2].Cnv_Level[1].Cnv1.Barcode_ID := 8;
   LCnv_Sys[2].Cnv_Level[2].Cnv1.Barcode_ID := 16;
   LCnv_Sys[2].Cnv_Level[3].Cnv1.Barcode_ID := 24;
   LCnv_Sys[2].Cnv_Level[4].Cnv1.Barcode_ID := 32;
   LCnv_Sys[2].Cnv_Level[5].Cnv1.Barcode_ID := 40;
   LCnv_Sys[2].Cnv_Level[6].Cnv1.Barcode_ID := 48;
   LCnv_Sys[2].Cnv_Level[7].Cnv1.Barcode_ID := 56;
   LCnv_Sys[2].Cnv_Level[8].Cnv1.Barcode_ID := 64;
   LCnv_Sys[3].Cnv_Level[1].Cnv1.Barcode_ID := 10;
   LCnv_Sys[3].Cnv_Level[2].Cnv1.Barcode_ID := 18;
   LCnv_Sys[3].Cnv_Level[3].Cnv1.Barcode_ID := 26;
   LCnv_Sys[3].Cnv_Level[4].Cnv1.Barcode_ID := 34;
   LCnv_Sys[3].Cnv_Level[5].Cnv1.Barcode_ID := 42;
   LCnv_Sys[3].Cnv_Level[6].Cnv1.Barcode_ID := 50;
   LCnv_Sys[3].Cnv_Level[7].Cnv1.Barcode_ID := 58;
   LCnv_Sys[3].Cnv_Level[8].Cnv1.Barcode_ID := 66;
   LCnv_Sys[4].Cnv_Level[1].Cnv1.Barcode_ID := 12;
   LCnv_Sys[4].Cnv_Level[2].Cnv1.Barcode_ID := 20;
   LCnv_Sys[4].Cnv_Level[3].Cnv1.Barcode_ID := 28;
   LCnv_Sys[4].Cnv_Level[4].Cnv1.Barcode_ID := 36;
   LCnv_Sys[4].Cnv_Level[5].Cnv1.Barcode_ID := 44;
   LCnv_Sys[4].Cnv_Level[6].Cnv1.Barcode_ID := 52;
   LCnv_Sys[4].Cnv_Level[7].Cnv1.Barcode_ID := 60;
   LCnv_Sys[4].Cnv_Level[8].Cnv1.Barcode_ID := 68;
   LCnv_Sys[5].Cnv_Level[1].Cnv1.Barcode_ID := 13;
   LCnv_Sys[5].Cnv_Level[2].Cnv1.Barcode_ID := 21;
   LCnv_Sys[5].Cnv_Level[3].Cnv1.Barcode_ID := 29;
   LCnv_Sys[5].Cnv_Level[4].Cnv1.Barcode_ID := 37;
   LCnv_Sys[5].Cnv_Level[5].Cnv1.Barcode_ID := 45;
   LCnv_Sys[5].Cnv_Level[6].Cnv1.Barcode_ID := 53;
   LCnv_Sys[5].Cnv_Level[7].Cnv1.Barcode_ID := 61;
   LCnv_Sys[5].Cnv_Level[8].Cnv1.Barcode_ID := 69;
   LCnv_Sys[1].Cnv_Level[1].Cnv1.Cnv_Level := 1;
   LCnv_Sys[1].Cnv_Level[2].Cnv1.Cnv_Level := 2;
   LCnv_Sys[1].Cnv_Level[3].Cnv1.Cnv_Level := 3;
   LCnv_Sys[1].Cnv_Level[4].Cnv1.Cnv_Level := 4;
   LCnv_Sys[1].Cnv_Level[5].Cnv1.Cnv_Level := 5;
   LCnv_Sys[1].Cnv_Level[6].Cnv1.Cnv_Level := 6;
   LCnv_Sys[1].Cnv_Level[7].Cnv1.Cnv_Level := 7;
   LCnv_Sys[1].Cnv_Level[8].Cnv1.Cnv_Level := 8;
   LCnv_Sys[2].Cnv_Level[1].Cnv1.Cnv_Level := 1;
   LCnv_Sys[2].Cnv_Level[2].Cnv1.Cnv_Level := 2;
   LCnv_Sys[2].Cnv_Level[3].Cnv1.Cnv_Level := 3;
   LCnv_Sys[2].Cnv_Level[4].Cnv1.Cnv_Level := 4;
   LCnv_Sys[2].Cnv_Level[5].Cnv1.Cnv_Level := 5;
   LCnv_Sys[2].Cnv_Level[6].Cnv1.Cnv_Level := 6;
   LCnv_Sys[2].Cnv_Level[7].Cnv1.Cnv_Level := 7;
   LCnv_Sys[2].Cnv_Level[8].Cnv1.Cnv_Level := 8;
   LCnv_Sys[3].Cnv_Level[1].Cnv1.Cnv_Level := 1;
   LCnv_Sys[3].Cnv_Level[2].Cnv1.Cnv_Level := 2;
   LCnv_Sys[3].Cnv_Level[3].Cnv1.Cnv_Level := 3;
   LCnv_Sys[3].Cnv_Level[4].Cnv1.Cnv_Level := 4;
   LCnv_Sys[3].Cnv_Level[5].Cnv1.Cnv_Level := 5;
   LCnv_Sys[3].Cnv_Level[6].Cnv1.Cnv_Level := 6;
   LCnv_Sys[3].Cnv_Level[7].Cnv1.Cnv_Level := 7;
   LCnv_Sys[3].Cnv_Level[8].Cnv1.Cnv_Level := 8;
   LCnv_Sys[4].Cnv_Level[1].Cnv1.Cnv_Level := 1;
   LCnv_Sys[4].Cnv_Level[2].Cnv1.Cnv_Level := 2;
   LCnv_Sys[4].Cnv_Level[3].Cnv1.Cnv_Level := 3;
   LCnv_Sys[4].Cnv_Level[4].Cnv1.Cnv_Level := 4;
   LCnv_Sys[4].Cnv_Level[5].Cnv1.Cnv_Level := 5;
   LCnv_Sys[4].Cnv_Level[6].Cnv1.Cnv_Level := 6;
   LCnv_Sys[4].Cnv_Level[7].Cnv1.Cnv_Level := 7;
   LCnv_Sys[4].Cnv_Level[8].Cnv1.Cnv_Level := 8;
   LCnv_Sys[5].Cnv_Level[1].Cnv1.Cnv_Level := 1;
   LCnv_Sys[5].Cnv_Level[2].Cnv1.Cnv_Level := 2;
   LCnv_Sys[5].Cnv_Level[3].Cnv1.Cnv_Level := 3;
   LCnv_Sys[5].Cnv_Level[4].Cnv1.Cnv_Level := 4;
   LCnv_Sys[5].Cnv_Level[5].Cnv1.Cnv_Level := 5;
   LCnv_Sys[5].Cnv_Level[6].Cnv1.Cnv_Level := 6;
   LCnv_Sys[5].Cnv_Level[7].Cnv1.Cnv_Level := 7;
   LCnv_Sys[5].Cnv_Level[8].Cnv1.Cnv_Level := 8;
   LCnv_Sys[1].Cnv_Level[1..8].Cnv1.TC_Time := 20;
   LCnv_Sys[2].Cnv_Level[1..8].Cnv1.TC_Time := 20;
   LCnv_Sys[3].Cnv_Level[1..8].Cnv1.TC_Time := 20;
   LCnv_Sys[4].Cnv_Level[1..8].Cnv1.TC_Time := 20;
   LCnv_Sys[5].Cnv_Level[1..8].Cnv1.TC_Time := 20;
   LCnv_Sys[1].Cnv_Level[1..8].Cnv1.Transfer_Time := 20;
   LCnv_Sys[2].Cnv_Level[1..8].Cnv1.Transfer_Time := 20;
   LCnv_Sys[3].Cnv_Level[1..8].Cnv1.Transfer_Time := 20;
   LCnv_Sys[4].Cnv_Level[1..3].Cnv1.Transfer_Time := 20;
   LCnv_Sys[4].Cnv_Level[4..8].Cnv1.Transfer_Time := 15;
   LCnv_Sys[5].Cnv_Level[1..8].Cnv1.Transfer_Time := 15;
   LCnv_Sys[1].Cnv_Level[1..8].Cnv1.Pallet_Align_Time := 20;
   LCnv_Sys[2].Cnv_Level[1..8].Cnv1.Pallet_Align_Time := 20;
   LCnv_Sys[3].Cnv_Level[1..8].Cnv1.Pallet_Align_Time := 20;
   LCnv_Sys[4].Cnv_Level[1..8].Cnv1.Pallet_Align_Time := 20;
   LCnv_Sys[5].Cnv_Level[1..8].Cnv1.Pallet_Align_Time := 20;
   LCnv_Sys[1].Cnv_Level[1..8].Cnv1.Slow_Speed := 11;
   LCnv_Sys[2].Cnv_Level[1..8].Cnv1.Slow_Speed := 11;
   LCnv_Sys[3].Cnv_Level[1..8].Cnv1.Slow_Speed := 11;
   LCnv_Sys[4].Cnv_Level[1..8].Cnv1.Slow_Speed := 11;
   LCnv_Sys[5].Cnv_Level[1..8].Cnv1.Slow_Speed := 11;
   LCnv_Sys[1].Cnv_Level[1..8].Cnv1.Full_Speed := 86;
   LCnv_Sys[2].Cnv_Level[1..8].Cnv1.Full_Speed := 86;
   LCnv_Sys[3].Cnv_Level[1..8].Cnv1.Full_Speed := 86;
   LCnv_Sys[4].Cnv_Level[1..8].Cnv1.Full_Speed := 86;
   LCnv_Sys[5].Cnv_Level[1..8].Cnv1.Full_Speed := 86;
   LCnv_Sys[1].Cnv_Level[1].Cnv1.Manual_Speed := 90;
   LCnv_Sys[1].Cnv_Level[2..8].Cnv1.Manual_Speed := 40;
   LCnv_Sys[2].Cnv_Level[1..8].Cnv1.Manual_Speed := 40;
   LCnv_Sys[3].Cnv_Level[1..8].Cnv1.Manual_Speed := 40;
   LCnv_Sys[4].Cnv_Level[1..8].Cnv1.Manual_Speed := 40;
   LCnv_Sys[5].Cnv_Level[1..8].Cnv1.Manual_Speed := 40;
   LCnv_Sys[1].Cnv_Level[1..8].Cnv1.Safety_stop_Timeout := 3000;
   LCnv_Sys[2].Cnv_Level[1..8].Cnv1.Safety_stop_Timeout := 3000;
   LCnv_Sys[3].Cnv_Level[1..8].Cnv1.Safety_stop_Timeout := 3000;
   LCnv_Sys[4].Cnv_Level[1..8].Cnv1.Safety_stop_Timeout := 3000;
   LCnv_Sys[5].Cnv_Level[1..8].Cnv1.Safety_stop_Timeout := 3000;
   LCnv_Sys[1].Cnv_Level[1..8].Cnv1.Timer_Check_Pallet_Time := 500;
   LCnv_Sys[2].Cnv_Level[1..8].Cnv1.Timer_Check_Pallet_Time := 500;
   LCnv_Sys[3].Cnv_Level[1..8].Cnv1.Timer_Check_Pallet_Time := 500;
   LCnv_Sys[4].Cnv_Level[1..8].Cnv1.Timer_Check_Pallet_Time := 500;
   LCnv_Sys[5].Cnv_Level[1..8].Cnv1.Timer_Check_Pallet_Time := 500;
   LCnv_Sys[1].Cnv_Level[1].Cnv1.G120_Hardware_ID := 527;
   LCnv_Sys[1].Cnv_Level[2].Cnv1.G120_Hardware_ID := 551;
   LCnv_Sys[1].Cnv_Level[3].Cnv1.G120_Hardware_ID := 569;
   LCnv_Sys[1].Cnv_Level[4].Cnv1.G120_Hardware_ID := 581;
   LCnv_Sys[1].Cnv_Level[5].Cnv1.G120_Hardware_ID := 593;
   LCnv_Sys[1].Cnv_Level[6].Cnv1.G120_Hardware_ID := 605;
   LCnv_Sys[1].Cnv_Level[7].Cnv1.G120_Hardware_ID := 726;
   LCnv_Sys[1].Cnv_Level[8].Cnv1.G120_Hardware_ID := 617;
   LCnv_Sys[2].Cnv_Level[1].Cnv1.G120_Hardware_ID := 980;
   LCnv_Sys[2].Cnv_Level[2].Cnv1.G120_Hardware_ID := 996;
   LCnv_Sys[2].Cnv_Level[3].Cnv1.G120_Hardware_ID := 1008;
   LCnv_Sys[2].Cnv_Level[4].Cnv1.G120_Hardware_ID := 1020;
   LCnv_Sys[2].Cnv_Level[5].Cnv1.G120_Hardware_ID := 1056;
   LCnv_Sys[2].Cnv_Level[6].Cnv1.G120_Hardware_ID := 1032;
   LCnv_Sys[2].Cnv_Level[7].Cnv1.G120_Hardware_ID := 1044;
   LCnv_Sys[2].Cnv_Level[8].Cnv1.G120_Hardware_ID := 1068;
   LCnv_Sys[3].Cnv_Level[1].Cnv1.G120_Hardware_ID := 1384;
   LCnv_Sys[3].Cnv_Level[2].Cnv1.G120_Hardware_ID := 1400;
   LCnv_Sys[3].Cnv_Level[3].Cnv1.G120_Hardware_ID := 1412;
   LCnv_Sys[3].Cnv_Level[4].Cnv1.G120_Hardware_ID := 1424;
   LCnv_Sys[3].Cnv_Level[5].Cnv1.G120_Hardware_ID := 1436;
   LCnv_Sys[3].Cnv_Level[6].Cnv1.G120_Hardware_ID := 1448;
   LCnv_Sys[3].Cnv_Level[7].Cnv1.G120_Hardware_ID := 1460;
   LCnv_Sys[3].Cnv_Level[8].Cnv1.G120_Hardware_ID := 1472;
   LCnv_Sys[4].Cnv_Level[1].Cnv1.G120_Hardware_ID := 1788;
   LCnv_Sys[4].Cnv_Level[2].Cnv1.G120_Hardware_ID := 1804;
   LCnv_Sys[4].Cnv_Level[3].Cnv1.G120_Hardware_ID := 1816;
   LCnv_Sys[4].Cnv_Level[4].Cnv1.G120_Hardware_ID := 1828;
   LCnv_Sys[4].Cnv_Level[5].Cnv1.G120_Hardware_ID := 1840;
   LCnv_Sys[4].Cnv_Level[6].Cnv1.G120_Hardware_ID := 1852;
   LCnv_Sys[4].Cnv_Level[7].Cnv1.G120_Hardware_ID := 1864;
   LCnv_Sys[4].Cnv_Level[8].Cnv1.G120_Hardware_ID := 1876;
   LCnv_Sys[5].Cnv_Level[1].Cnv1.G120_Hardware_ID := 2096;
   LCnv_Sys[5].Cnv_Level[2].Cnv1.G120_Hardware_ID := 2112;
   LCnv_Sys[5].Cnv_Level[3].Cnv1.G120_Hardware_ID := 2124;
   LCnv_Sys[5].Cnv_Level[4].Cnv1.G120_Hardware_ID := 2136;
   LCnv_Sys[5].Cnv_Level[5].Cnv1.G120_Hardware_ID := 2148;
   LCnv_Sys[5].Cnv_Level[6].Cnv1.G120_Hardware_ID := 2160;
   LCnv_Sys[5].Cnv_Level[7].Cnv1.G120_Hardware_ID := 2172;
   LCnv_Sys[5].Cnv_Level[8].Cnv1.G120_Hardware_ID := 2184;
   LCnv_Sys[1].Cnv_Level[1].Cnv2.ID := 110101;
   LCnv_Sys[1].Cnv_Level[2].Cnv2.ID := 110201;
   LCnv_Sys[1].Cnv_Level[3].Cnv2.ID := 110301;
   LCnv_Sys[1].Cnv_Level[4].Cnv2.ID := 110401;
   LCnv_Sys[1].Cnv_Level[5].Cnv2.ID := 110501;
   LCnv_Sys[1].Cnv_Level[6].Cnv2.ID := 110601;
   LCnv_Sys[1].Cnv_Level[7].Cnv2.ID := 110701;
   LCnv_Sys[1].Cnv_Level[8].Cnv2.ID := 110801;
   LCnv_Sys[2].Cnv_Level[1].Cnv2.ID := 110102;
   LCnv_Sys[2].Cnv_Level[2].Cnv2.ID := 110202;
   LCnv_Sys[2].Cnv_Level[3].Cnv2.ID := 110302;
   LCnv_Sys[2].Cnv_Level[4].Cnv2.ID := 110402;
   LCnv_Sys[2].Cnv_Level[5].Cnv2.ID := 110502;
   LCnv_Sys[2].Cnv_Level[6].Cnv2.ID := 110602;
   LCnv_Sys[2].Cnv_Level[7].Cnv2.ID := 110702;
   LCnv_Sys[2].Cnv_Level[8].Cnv2.ID := 110802;
   LCnv_Sys[3].Cnv_Level[1].Cnv2.ID := 110103;
   LCnv_Sys[3].Cnv_Level[2].Cnv2.ID := 110203;
   LCnv_Sys[3].Cnv_Level[3].Cnv2.ID := 110303;
   LCnv_Sys[3].Cnv_Level[4].Cnv2.ID := 110403;
   LCnv_Sys[3].Cnv_Level[5].Cnv2.ID := 110503;
   LCnv_Sys[3].Cnv_Level[6].Cnv2.ID := 110603;
   LCnv_Sys[3].Cnv_Level[7].Cnv2.ID := 110703;
   LCnv_Sys[3].Cnv_Level[8].Cnv2.ID := 110803;
   LCnv_Sys[4].Cnv_Level[1].Cnv2.ID := 110104;
   LCnv_Sys[4].Cnv_Level[2].Cnv2.ID := 110204;
   LCnv_Sys[4].Cnv_Level[3].Cnv2.ID := 110304;
   LCnv_Sys[4].Cnv_Level[4].Cnv2.ID := 110404;
   LCnv_Sys[4].Cnv_Level[5].Cnv2.ID := 110504;
   LCnv_Sys[4].Cnv_Level[6].Cnv2.ID := 110604;
   LCnv_Sys[4].Cnv_Level[7].Cnv2.ID := 110704;
   LCnv_Sys[4].Cnv_Level[8].Cnv2.ID := 110804;
   LCnv_Sys[5].Cnv_Level[1].Cnv2.ID := 110105;
   LCnv_Sys[5].Cnv_Level[2].Cnv2.ID := 110205;
   LCnv_Sys[5].Cnv_Level[3].Cnv2.ID := 110305;
   LCnv_Sys[5].Cnv_Level[4].Cnv2.ID := 110405;
   LCnv_Sys[5].Cnv_Level[5].Cnv2.ID := 110505;
   LCnv_Sys[5].Cnv_Level[6].Cnv2.ID := 110605;
   LCnv_Sys[5].Cnv_Level[7].Cnv2.ID := 110705;
   LCnv_Sys[5].Cnv_Level[8].Cnv2.ID := 110805;
   LCnv_Sys[1].Cnv_Level[1].Cnv2.Barcode_ID := 7;
   LCnv_Sys[1].Cnv_Level[2].Cnv2.Barcode_ID := 15;
   LCnv_Sys[1].Cnv_Level[3].Cnv2.Barcode_ID := 23;
   LCnv_Sys[1].Cnv_Level[4].Cnv2.Barcode_ID := 31;
   LCnv_Sys[1].Cnv_Level[5].Cnv2.Barcode_ID := 39;
   LCnv_Sys[1].Cnv_Level[6].Cnv2.Barcode_ID := 47;
   LCnv_Sys[1].Cnv_Level[7].Cnv2.Barcode_ID := 55;
   LCnv_Sys[1].Cnv_Level[8].Cnv2.Barcode_ID := 63;
   LCnv_Sys[2].Cnv_Level[1].Cnv2.Barcode_ID := 9;
   LCnv_Sys[2].Cnv_Level[2].Cnv2.Barcode_ID := 17;
   LCnv_Sys[2].Cnv_Level[3].Cnv2.Barcode_ID := 25;
   LCnv_Sys[2].Cnv_Level[4].Cnv2.Barcode_ID := 33;
   LCnv_Sys[2].Cnv_Level[5].Cnv2.Barcode_ID := 41;
   LCnv_Sys[2].Cnv_Level[6].Cnv2.Barcode_ID := 49;
   LCnv_Sys[2].Cnv_Level[7].Cnv2.Barcode_ID := 57;
   LCnv_Sys[2].Cnv_Level[8].Cnv2.Barcode_ID := 65;
   LCnv_Sys[3].Cnv_Level[1].Cnv2.Barcode_ID := 11;
   LCnv_Sys[3].Cnv_Level[2].Cnv2.Barcode_ID := 19;
   LCnv_Sys[3].Cnv_Level[3].Cnv2.Barcode_ID := 27;
   LCnv_Sys[3].Cnv_Level[4].Cnv2.Barcode_ID := 35;
   LCnv_Sys[3].Cnv_Level[5].Cnv2.Barcode_ID := 43;
   LCnv_Sys[3].Cnv_Level[6].Cnv2.Barcode_ID := 51;
   LCnv_Sys[3].Cnv_Level[7].Cnv2.Barcode_ID := 59;
   LCnv_Sys[3].Cnv_Level[8].Cnv2.Barcode_ID := 67;
   LCnv_Sys[4].Cnv_Level[1..8].Cnv2.Barcode_ID := 0;
   LCnv_Sys[5].Cnv_Level[1..8].Cnv2.Barcode_ID := 0;
   LCnv_Sys[1].Cnv_Level[1].Cnv2.Cnv_Level := 1;
   LCnv_Sys[1].Cnv_Level[2].Cnv2.Cnv_Level := 2;
   LCnv_Sys[1].Cnv_Level[3].Cnv2.Cnv_Level := 3;
   LCnv_Sys[1].Cnv_Level[4].Cnv2.Cnv_Level := 4;
   LCnv_Sys[1].Cnv_Level[5].Cnv2.Cnv_Level := 5;
   LCnv_Sys[1].Cnv_Level[6].Cnv2.Cnv_Level := 6;
   LCnv_Sys[1].Cnv_Level[7].Cnv2.Cnv_Level := 7;
   LCnv_Sys[1].Cnv_Level[8].Cnv2.Cnv_Level := 8;
   LCnv_Sys[2].Cnv_Level[1].Cnv2.Cnv_Level := 1;
   LCnv_Sys[2].Cnv_Level[2].Cnv2.Cnv_Level := 2;
   LCnv_Sys[2].Cnv_Level[3].Cnv2.Cnv_Level := 3;
   LCnv_Sys[2].Cnv_Level[4].Cnv2.Cnv_Level := 4;
   LCnv_Sys[2].Cnv_Level[5].Cnv2.Cnv_Level := 5;
   LCnv_Sys[2].Cnv_Level[6].Cnv2.Cnv_Level := 6;
   LCnv_Sys[2].Cnv_Level[7].Cnv2.Cnv_Level := 7;
   LCnv_Sys[2].Cnv_Level[8].Cnv2.Cnv_Level := 8;
   LCnv_Sys[3].Cnv_Level[1].Cnv2.Cnv_Level := 1;
   LCnv_Sys[3].Cnv_Level[2].Cnv2.Cnv_Level := 2;
   LCnv_Sys[3].Cnv_Level[3].Cnv2.Cnv_Level := 3;
   LCnv_Sys[3].Cnv_Level[4].Cnv2.Cnv_Level := 4;
   LCnv_Sys[3].Cnv_Level[5].Cnv2.Cnv_Level := 5;
   LCnv_Sys[3].Cnv_Level[6].Cnv2.Cnv_Level := 6;
   LCnv_Sys[3].Cnv_Level[7].Cnv2.Cnv_Level := 7;
   LCnv_Sys[3].Cnv_Level[8].Cnv2.Cnv_Level := 8;
   LCnv_Sys[4].Cnv_Level[1..8].Cnv2.Cnv_Level := 1;
   LCnv_Sys[5].Cnv_Level[1..8].Cnv2.Cnv_Level := 1;
   LCnv_Sys[1].Cnv_Level[1..8].Cnv2.TC_Time := 20;
   LCnv_Sys[2].Cnv_Level[1..8].Cnv2.TC_Time := 20;
   LCnv_Sys[3].Cnv_Level[1..8].Cnv2.TC_Time := 20;
   LCnv_Sys[4].Cnv_Level[1..8].Cnv2.TC_Time := 20;
   LCnv_Sys[5].Cnv_Level[1..8].Cnv2.TC_Time := 20;
   LCnv_Sys[1].Cnv_Level[1..8].Cnv2.Transfer_Time := 20;
   LCnv_Sys[2].Cnv_Level[1..8].Cnv2.Transfer_Time := 20;
   LCnv_Sys[3].Cnv_Level[1..8].Cnv2.Transfer_Time := 20;
   LCnv_Sys[4].Cnv_Level[1..2].Cnv2.Transfer_Time := 20;
   LCnv_Sys[4].Cnv_Level[3..8].Cnv2.Transfer_Time := 15;
   LCnv_Sys[5].Cnv_Level[1..8].Cnv2.Transfer_Time := 15;
   LCnv_Sys[1].Cnv_Level[1..8].Cnv2.Pallet_Align_Time := 20;
   LCnv_Sys[2].Cnv_Level[1..8].Cnv2.Pallet_Align_Time := 20;
   LCnv_Sys[3].Cnv_Level[1..8].Cnv2.Pallet_Align_Time := 20;
   LCnv_Sys[4].Cnv_Level[1..8].Cnv2.Pallet_Align_Time := 20;
   LCnv_Sys[5].Cnv_Level[1..8].Cnv2.Pallet_Align_Time := 20;
   LCnv_Sys[1].Cnv_Level[1..8].Cnv2.Slow_Speed := 11;
   LCnv_Sys[2].Cnv_Level[1..8].Cnv2.Slow_Speed := 11;
   LCnv_Sys[3].Cnv_Level[1..8].Cnv2.Slow_Speed := 11;
   LCnv_Sys[4].Cnv_Level[1..8].Cnv2.Slow_Speed := 10;
   LCnv_Sys[5].Cnv_Level[1..8].Cnv2.Slow_Speed := 10;
   LCnv_Sys[1].Cnv_Level[1..8].Cnv2.Full_Speed := 86;
   LCnv_Sys[2].Cnv_Level[1..8].Cnv2.Full_Speed := 86;
   LCnv_Sys[3].Cnv_Level[1..8].Cnv2.Full_Speed := 86;
   LCnv_Sys[4].Cnv_Level[1..8].Cnv2.Full_Speed := 86;
   LCnv_Sys[5].Cnv_Level[1..8].Cnv2.Full_Speed := 86;
   LCnv_Sys[1].Cnv_Level[1..8].Cnv2.Manual_Speed := 40;
   LCnv_Sys[2].Cnv_Level[1..8].Cnv2.Manual_Speed := 40;
   LCnv_Sys[3].Cnv_Level[1..8].Cnv2.Manual_Speed := 40;
   LCnv_Sys[4].Cnv_Level[1..8].Cnv2.Manual_Speed := 40;
   LCnv_Sys[5].Cnv_Level[1..8].Cnv2.Manual_Speed := 40;
   LCnv_Sys[1].Cnv_Level[1..8].Cnv2.Safety_stop_Timeout := 3000;
   LCnv_Sys[2].Cnv_Level[1..8].Cnv2.Safety_stop_Timeout := 3000;
   LCnv_Sys[3].Cnv_Level[1..8].Cnv2.Safety_stop_Timeout := 3000;
   LCnv_Sys[4].Cnv_Level[1..4].Cnv2.Safety_stop_Timeout := 3000;
   LCnv_Sys[4].Cnv_Level[5..8].Cnv2.Safety_stop_Timeout := 20;
   LCnv_Sys[5].Cnv_Level[1..8].Cnv2.Safety_stop_Timeout := 20;
   LCnv_Sys[1].Cnv_Level[1..8].Cnv2.Timer_Check_Pallet_Time := 500;
   LCnv_Sys[2].Cnv_Level[1..8].Cnv2.Timer_Check_Pallet_Time := 500;
   LCnv_Sys[3].Cnv_Level[1..8].Cnv2.Timer_Check_Pallet_Time := 500;
   LCnv_Sys[1].Cnv_Level[1].Cnv2.G120_Hardware_ID := 629;
   LCnv_Sys[1].Cnv_Level[2].Cnv2.G120_Hardware_ID := 641;
   LCnv_Sys[1].Cnv_Level[3].Cnv2.G120_Hardware_ID := 653;
   LCnv_Sys[1].Cnv_Level[4].Cnv2.G120_Hardware_ID := 665;
   LCnv_Sys[1].Cnv_Level[5].Cnv2.G120_Hardware_ID := 678;
   LCnv_Sys[1].Cnv_Level[6].Cnv2.G120_Hardware_ID := 690;
   LCnv_Sys[1].Cnv_Level[7].Cnv2.G120_Hardware_ID := 702;
   LCnv_Sys[1].Cnv_Level[8].Cnv2.G120_Hardware_ID := 714;
   LCnv_Sys[2].Cnv_Level[1].Cnv2.G120_Hardware_ID := 1080;
   LCnv_Sys[2].Cnv_Level[2].Cnv2.G120_Hardware_ID := 1092;
   LCnv_Sys[2].Cnv_Level[3].Cnv2.G120_Hardware_ID := 1104;
   LCnv_Sys[2].Cnv_Level[4].Cnv2.G120_Hardware_ID := 1116;
   LCnv_Sys[2].Cnv_Level[5].Cnv2.G120_Hardware_ID := 1128;
   LCnv_Sys[2].Cnv_Level[6].Cnv2.G120_Hardware_ID := 1140;
   LCnv_Sys[2].Cnv_Level[7].Cnv2.G120_Hardware_ID := 1152;
   LCnv_Sys[2].Cnv_Level[8].Cnv2.G120_Hardware_ID := 1164;
   LCnv_Sys[3].Cnv_Level[1].Cnv2.G120_Hardware_ID := 1484;
   LCnv_Sys[3].Cnv_Level[2].Cnv2.G120_Hardware_ID := 1496;
   LCnv_Sys[3].Cnv_Level[3].Cnv2.G120_Hardware_ID := 1508;
   LCnv_Sys[3].Cnv_Level[4].Cnv2.G120_Hardware_ID := 1520;
   LCnv_Sys[3].Cnv_Level[5].Cnv2.G120_Hardware_ID := 1532;
   LCnv_Sys[3].Cnv_Level[6].Cnv2.G120_Hardware_ID := 1544;
   LCnv_Sys[3].Cnv_Level[7].Cnv2.G120_Hardware_ID := 1556;
   LCnv_Sys[3].Cnv_Level[8].Cnv2.G120_Hardware_ID := 1568;
   LCnv_Sys[4].Cnv_Level[1..8].Cnv2.G120_Hardware_ID := 0;
   LCnv_Sys[5].Cnv_Level[1..8].Cnv2.G120_Hardware_ID := 0;
   Shuttle_MQTT.MQTT_Con_Params.hwId := 0;
   Shuttle_MQTT.MQTT_Con_Params.connId := 16#0001;
   Shuttle_MQTT.MQTT_Con_Params.broker := '10.44.116.8';
   Shuttle_MQTT.MQTT_Con_Params.port := 1883;
   Shuttle_MQTT.MQTT_Con_Params.tls.enableTls := FALSE;
   Shuttle_MQTT.MQTT_Con_Params.tls.validateServerIdentity := FALSE;
   Shuttle_MQTT.MQTT_Con_Params.tls.brokerCert := 0;
   Shuttle_MQTT.MQTT_Con_Params.tls.clientCert := 0;
   Shuttle_MQTT.MQTT_Con_Params.keepAlive := 60;
   Shuttle_MQTT.Client_ID := WSTRING#'PLC_1';
   Shuttle_MQTT.Username := WSTRING#'';
   Shuttle_MQTT.Password := WSTRING#'';
   Shuttle_MQTT.Timeout := 0;
   Shuttle_MQTT.QoS := 0;
   Shuttle_MQTT.Retain := TRUE;
   Shuttle_MQTT.Will_Topic := WSTRING#'';
   Shuttle_MQTT.Will_Msg_Length := 0;
   Shuttle_MQTT.Will_Msg_Payload[1..128] := 16#00;
   System.VTD_Count := 5;
   System.Level_Count := 8;
   System.Cnv_Count := 95;
   System.Shuttle_Count := 23;
   System.Shuttle_Interlock_Timeout := 999;
END_DATA_BLOCK

DATA_BLOCK "Shuttle_MQTT_DB"   // DB75
{ S7_Optimized_Access := 'TRUE' }
VERSION : 0.1
// stored: AutoNumber true, DBAccessibleFromOPCUA true, IsOnlyStoredInLoadMemory false, IsRetainMemResEnabled false, IsWriteProtectedInAS false, MemoryReserve 100
   VAR
      Shuttle_MQTT : Array[1..24] of "MQTT_Interface";
   END_VAR
BEGIN
END_DATA_BLOCK

DATA_BLOCK "TCP_IP_Shuttle_DB_1"   // DB391
{ S7_Optimized_Access := 'TRUE' }
VERSION : 0.1
// stored: AutoNumber true, DBAccessibleFromOPCUA true, IsOnlyStoredInLoadMemory false, IsRetainMemResEnabled false, IsWriteProtectedInAS false, MemoryReserve 100
   VAR
      enable : Bool := TRUE;
      send : Bool;
      sendDataLength : UDInt := 0;
      receiveDataLength : UDInt := 16#FFFF_FFFF;
   END_VAR
   VAR RETAIN
      tcpConfig : "LCom_typeConfig";
   END_VAR
   VAR
      tcpDiagnostics { S7_SetPoint := 'True'} : "LCom_typeDiagnostics";
      sendBuffer { S7_SetPoint := 'True'} : Array[0..59] of Byte;
      SendBufferSize : UInt := 60;
      receiveBuffer : Array[0..27] of Byte;
      receiveBufferSize : UInt := 28;
      connected : Bool;
      sending : Bool;
      dataReceived : Bool;
      receivedDataLength : UDInt;
      busy : Bool;
      error : Bool;
      status : Word;
   END_VAR
BEGIN
   tcpConfig.connection.interfaceID := 65164;
   tcpConfig.connection.connectionID := 101;
   tcpConfig.connection.comService := 1;
   tcpConfig.connection.isClient := False;
   tcpConfig.connection.connectType := 1;
   tcpConfig.connection.localPort := 4001;
   tcpConfig.connection.partnerPort := 4001;
   tcpConfig.connection.partnerIP.ADDR[1] := 10;
   tcpConfig.connection.partnerIP.ADDR[2] := 0;
   tcpConfig.connection.partnerIP.ADDR[3] := 34;
   tcpConfig.connection.partnerIP.ADDR[4] := 211;
   tcpConfig.connection.acceptUnknownPartner := TRUE;
   tcpConfig.connection.lifeSignCycleTime := T#1s;
   // sendBuffer[0] : STX
   // sendBuffer[1] : Size
   // sendBuffer[2] : Type
   // sendBuffer[3] : Request ID 1
   // sendBuffer[4] : Request ID 2
   // sendBuffer[5] : PID 1
   // sendBuffer[6] : PID 2
   // sendBuffer[7] : PID 3
   // sendBuffer[8] : PID 4
   // sendBuffer[9] : DID 1
   // sendBuffer[10] : DID 2
   // sendBuffer[11] : DID 3
   // sendBuffer[12] : DID 4
   // sendBuffer[13] : Distance remaining 1
   // sendBuffer[14] : Distance remaining 2
   // sendBuffer[15] : X
   // sendBuffer[16] : X
   // sendBuffer[17] : X
   // sendBuffer[18] : X
   // sendBuffer[19] : Y
   // sendBuffer[20] : Y
   // sendBuffer[21] : Y
   // sendBuffer[22] : Y
   // sendBuffer[23] : Floor
   // sendBuffer[24] : Mode
   // sendBuffer[25] : State
   // sendBuffer[26] : Load State
   // sendBuffer[27] : E1
   // sendBuffer[28] : E1
   // sendBuffer[29] : E2
   // sendBuffer[30] : E2
   // sendBuffer[31] : E3
   // sendBuffer[32] : E3
   // sendBuffer[33] : E4
   // sendBuffer[34] : E4
   // sendBuffer[35] : E5
   // sendBuffer[36] : E5
   // sendBuffer[37] : E6
   // sendBuffer[38] : E6
   // sendBuffer[39] : I1
   // sendBuffer[40] : I1
   // sendBuffer[41] : Q1
   // sendBuffer[42] : Q1
   // sendBuffer[43] : Barcode 1
   // sendBuffer[44] : Barcode 2
   // sendBuffer[45] : Barcode 3
   // sendBuffer[46] : Barcode 4
   // sendBuffer[47] : Pallet Type
   // sendBuffer[48] : Energy Level
   // sendBuffer[49] : Battery Voltage
   // sendBuffer[50] : Battery Voltage
   // sendBuffer[51] : Paused
   // sendBuffer[52] : Last order 1
   // sendBuffer[53] : Last order 2
   // sendBuffer[54] : Current order 1
   // sendBuffer[55] : Current order 2
   // sendBuffer[56] : Last finished 1
   // sendBuffer[57] : Last Finished 2
   // sendBuffer[58] : CS
   // sendBuffer[59] : ETX
   // receiveBuffer[0] : STX
   // receiveBuffer[1] : Size (length of payload)
   // receiveBuffer[2] : Type
   // receiveBuffer[3] : Request ID 1
   // receiveBuffer[4] : Request ID 2
END_DATA_BLOCK

DATA_BLOCK "TCP_IP_Shuttle_DB_10"   // DB384
{ S7_Optimized_Access := 'TRUE' }
VERSION : 0.1
// stored: AutoNumber true, DBAccessibleFromOPCUA true, IsOnlyStoredInLoadMemory false, IsRetainMemResEnabled false, IsWriteProtectedInAS false, MemoryReserve 100
   VAR
      enable : Bool := TRUE;
      send : Bool;
      sendDataLength : UDInt := 0;
      receiveDataLength : UDInt := 16#FFFF_FFFF;
   END_VAR
   VAR RETAIN
      tcpConfig : "LCom_typeConfig";
   END_VAR
   VAR
      tcpDiagnostics { S7_SetPoint := 'True'} : "LCom_typeDiagnostics";
      sendBuffer { S7_SetPoint := 'True'} : Array[0..59] of Byte;
      SendBufferSize : UInt := 60;
      receiveBuffer : Array[0..27] of Byte;
      receiveBufferSize : UInt := 28;
      connected : Bool;
      sending : Bool;
      dataReceived : Bool;
      receivedDataLength : UDInt;
      busy : Bool;
      error : Bool;
      status : Word;
   END_VAR
BEGIN
   tcpConfig.connection.interfaceID := 65164;
   tcpConfig.connection.connectionID := 110;
   tcpConfig.connection.comService := 1;
   tcpConfig.connection.isClient := False;
   tcpConfig.connection.connectType := 1;
   tcpConfig.connection.localPort := 4010;
   tcpConfig.connection.partnerPort := 4010;
   tcpConfig.connection.partnerIP.ADDR[1] := 10;
   tcpConfig.connection.partnerIP.ADDR[2] := 0;
   tcpConfig.connection.partnerIP.ADDR[3] := 34;
   tcpConfig.connection.partnerIP.ADDR[4] := 220;
   tcpConfig.connection.acceptUnknownPartner := TRUE;
   tcpConfig.connection.lifeSignCycleTime := T#1s;
   // sendBuffer[0] : STX
   // sendBuffer[1] : Size
   // sendBuffer[2] : Type
   // sendBuffer[3] : Request ID 1
   // sendBuffer[4] : Request ID 2
   // sendBuffer[5] : PID 1
   // sendBuffer[6] : PID 2
   // sendBuffer[7] : PID 3
   // sendBuffer[8] : PID 4
   // sendBuffer[9] : DID 1
   // sendBuffer[10] : DID 2
   // sendBuffer[11] : DID 3
   // sendBuffer[12] : DID 4
   // sendBuffer[13] : Distance remaining 1
   // sendBuffer[14] : Distance remaining 2
   // sendBuffer[15] : X
   // sendBuffer[16] : X
   // sendBuffer[17] : X
   // sendBuffer[18] : X
   // sendBuffer[19] : Y
   // sendBuffer[20] : Y
   // sendBuffer[21] : Y
   // sendBuffer[22] : Y
   // sendBuffer[23] : Floor
   // sendBuffer[24] : Mode
   // sendBuffer[25] : State
   // sendBuffer[26] : Load State
   // sendBuffer[27] : E1
   // sendBuffer[28] : E1
   // sendBuffer[29] : E2
   // sendBuffer[30] : E2
   // sendBuffer[31] : E3
   // sendBuffer[32] : E3
   // sendBuffer[33] : E4
   // sendBuffer[34] : E4
   // sendBuffer[35] : E5
   // sendBuffer[36] : E5
   // sendBuffer[37] : E6
   // sendBuffer[38] : E6
   // sendBuffer[39] : I1
   // sendBuffer[40] : I1
   // sendBuffer[41] : Q1
   // sendBuffer[42] : Q1
   // sendBuffer[43] : Barcode 1
   // sendBuffer[44] : Barcode 2
   // sendBuffer[45] : Barcode 3
   // sendBuffer[46] : Barcode 4
   // sendBuffer[47] : Pallet Type
   // sendBuffer[48] : Energy Level
   // sendBuffer[49] : Battery Voltage
   // sendBuffer[50] : Battery Voltage
   // sendBuffer[51] : Paused
   // sendBuffer[52] : Last order 1
   // sendBuffer[53] : Last order 2
   // sendBuffer[54] : Current order 1
   // sendBuffer[55] : Current order 2
   // sendBuffer[56] : Last finished 1
   // sendBuffer[57] : Last Finished 2
   // sendBuffer[58] : CS
   // sendBuffer[59] : ETX
   // receiveBuffer[0] : STX
   // receiveBuffer[1] : Size (length of payload)
   // receiveBuffer[2] : Type
   // receiveBuffer[3] : Request ID 1
   // receiveBuffer[4] : Request ID 2
END_DATA_BLOCK

DATA_BLOCK "TCP_IP_Shuttle_DB_11"   // DB385
{ S7_Optimized_Access := 'TRUE' }
VERSION : 0.1
// stored: AutoNumber true, DBAccessibleFromOPCUA true, IsOnlyStoredInLoadMemory false, IsRetainMemResEnabled false, IsWriteProtectedInAS false, MemoryReserve 100
   VAR
      enable : Bool := TRUE;
      send : Bool;
      sendDataLength : UDInt := 0;
      receiveDataLength : UDInt := 16#FFFF_FFFF;
   END_VAR
   VAR RETAIN
      tcpConfig : "LCom_typeConfig";
   END_VAR
   VAR
      tcpDiagnostics { S7_SetPoint := 'True'} : "LCom_typeDiagnostics";
      sendBuffer { S7_SetPoint := 'True'} : Array[0..59] of Byte;
      SendBufferSize : UInt := 60;
      receiveBuffer : Array[0..27] of Byte;
      receiveBufferSize : UInt := 28;
      connected : Bool;
      sending : Bool;
      dataReceived : Bool;
      receivedDataLength : UDInt;
      busy : Bool;
      error : Bool;
      status : Word;
   END_VAR
BEGIN
   tcpConfig.connection.interfaceID := 65164;
   tcpConfig.connection.connectionID := 111;
   tcpConfig.connection.comService := 1;
   tcpConfig.connection.isClient := False;
   tcpConfig.connection.connectType := 1;
   tcpConfig.connection.localPort := 4011;
   tcpConfig.connection.partnerPort := 4011;
   tcpConfig.connection.partnerIP.ADDR[1] := 10;
   tcpConfig.connection.partnerIP.ADDR[2] := 0;
   tcpConfig.connection.partnerIP.ADDR[3] := 34;
   tcpConfig.connection.partnerIP.ADDR[4] := 221;
   tcpConfig.connection.acceptUnknownPartner := TRUE;
   tcpConfig.connection.lifeSignCycleTime := T#1s;
   // sendBuffer[0] : STX
   // sendBuffer[1] : Size
   // sendBuffer[2] : Type
   // sendBuffer[3] : Request ID 1
   // sendBuffer[4] : Request ID 2
   // sendBuffer[5] : PID 1
   // sendBuffer[6] : PID 2
   // sendBuffer[7] : PID 3
   // sendBuffer[8] : PID 4
   // sendBuffer[9] : DID 1
   // sendBuffer[10] : DID 2
   // sendBuffer[11] : DID 3
   // sendBuffer[12] : DID 4
   // sendBuffer[13] : Distance remaining 1
   // sendBuffer[14] : Distance remaining 2
   // sendBuffer[15] : X
   // sendBuffer[16] : X
   // sendBuffer[17] : X
   // sendBuffer[18] : X
   // sendBuffer[19] : Y
   // sendBuffer[20] : Y
   // sendBuffer[21] : Y
   // sendBuffer[22] : Y
   // sendBuffer[23] : Floor
   // sendBuffer[24] : Mode
   // sendBuffer[25] : State
   // sendBuffer[26] : Load State
   // sendBuffer[27] : E1
   // sendBuffer[28] : E1
   // sendBuffer[29] : E2
   // sendBuffer[30] : E2
   // sendBuffer[31] : E3
   // sendBuffer[32] : E3
   // sendBuffer[33] : E4
   // sendBuffer[34] : E4
   // sendBuffer[35] : E5
   // sendBuffer[36] : E5
   // sendBuffer[37] : E6
   // sendBuffer[38] : E6
   // sendBuffer[39] : I1
   // sendBuffer[40] : I1
   // sendBuffer[41] : Q1
   // sendBuffer[42] : Q1
   // sendBuffer[43] : Barcode 1
   // sendBuffer[44] : Barcode 2
   // sendBuffer[45] : Barcode 3
   // sendBuffer[46] : Barcode 4
   // sendBuffer[47] : Pallet Type
   // sendBuffer[48] : Energy Level
   // sendBuffer[49] : Battery Voltage
   // sendBuffer[50] : Battery Voltage
   // sendBuffer[51] : Paused
   // sendBuffer[52] : Last order 1
   // sendBuffer[53] : Last order 2
   // sendBuffer[54] : Current order 1
   // sendBuffer[55] : Current order 2
   // sendBuffer[56] : Last finished 1
   // sendBuffer[57] : Last Finished 2
   // sendBuffer[58] : CS
   // sendBuffer[59] : ETX
   // receiveBuffer[0] : STX
   // receiveBuffer[1] : Size (length of payload)
   // receiveBuffer[2] : Type
   // receiveBuffer[3] : Request ID 1
   // receiveBuffer[4] : Request ID 2
END_DATA_BLOCK

DATA_BLOCK "TCP_IP_Shuttle_DB_12"   // DB386
{ S7_Optimized_Access := 'TRUE' }
VERSION : 0.1
// stored: AutoNumber true, DBAccessibleFromOPCUA true, IsOnlyStoredInLoadMemory false, IsRetainMemResEnabled false, IsWriteProtectedInAS false, MemoryReserve 100
   VAR
      enable : Bool := TRUE;
      send : Bool;
      sendDataLength : UDInt := 0;
      receiveDataLength : UDInt := 16#FFFF_FFFF;
   END_VAR
   VAR RETAIN
      tcpConfig : "LCom_typeConfig";
   END_VAR
   VAR
      tcpDiagnostics { S7_SetPoint := 'True'} : "LCom_typeDiagnostics";
      sendBuffer { S7_SetPoint := 'True'} : Array[0..59] of Byte;
      SendBufferSize : UInt := 60;
      receiveBuffer : Array[0..27] of Byte;
      receiveBufferSize : UInt := 28;
      connected : Bool;
      sending : Bool;
      dataReceived : Bool;
      receivedDataLength : UDInt;
      busy : Bool;
      error : Bool;
      status : Word;
   END_VAR
BEGIN
   tcpConfig.connection.interfaceID := 65164;
   tcpConfig.connection.connectionID := 112;
   tcpConfig.connection.comService := 1;
   tcpConfig.connection.isClient := False;
   tcpConfig.connection.connectType := 1;
   tcpConfig.connection.localPort := 4012;
   tcpConfig.connection.partnerPort := 4012;
   tcpConfig.connection.partnerIP.ADDR[1] := 10;
   tcpConfig.connection.partnerIP.ADDR[2] := 0;
   tcpConfig.connection.partnerIP.ADDR[3] := 34;
   tcpConfig.connection.partnerIP.ADDR[4] := 222;
   tcpConfig.connection.acceptUnknownPartner := TRUE;
   tcpConfig.connection.lifeSignCycleTime := T#1s;
   // sendBuffer[0] : STX
   // sendBuffer[1] : Size
   // sendBuffer[2] : Type
   // sendBuffer[3] : Request ID 1
   // sendBuffer[4] : Request ID 2
   // sendBuffer[5] : PID 1
   // sendBuffer[6] : PID 2
   // sendBuffer[7] : PID 3
   // sendBuffer[8] : PID 4
   // sendBuffer[9] : DID 1
   // sendBuffer[10] : DID 2
   // sendBuffer[11] : DID 3
   // sendBuffer[12] : DID 4
   // sendBuffer[13] : Distance remaining 1
   // sendBuffer[14] : Distance remaining 2
   // sendBuffer[15] : X
   // sendBuffer[16] : X
   // sendBuffer[17] : X
   // sendBuffer[18] : X
   // sendBuffer[19] : Y
   // sendBuffer[20] : Y
   // sendBuffer[21] : Y
   // sendBuffer[22] : Y
   // sendBuffer[23] : Floor
   // sendBuffer[24] : Mode
   // sendBuffer[25] : State
   // sendBuffer[26] : Load State
   // sendBuffer[27] : E1
   // sendBuffer[28] : E1
   // sendBuffer[29] : E2
   // sendBuffer[30] : E2
   // sendBuffer[31] : E3
   // sendBuffer[32] : E3
   // sendBuffer[33] : E4
   // sendBuffer[34] : E4
   // sendBuffer[35] : E5
   // sendBuffer[36] : E5
   // sendBuffer[37] : E6
   // sendBuffer[38] : E6
   // sendBuffer[39] : I1
   // sendBuffer[40] : I1
   // sendBuffer[41] : Q1
   // sendBuffer[42] : Q1
   // sendBuffer[43] : Barcode 1
   // sendBuffer[44] : Barcode 2
   // sendBuffer[45] : Barcode 3
   // sendBuffer[46] : Barcode 4
   // sendBuffer[47] : Pallet Type
   // sendBuffer[48] : Energy Level
   // sendBuffer[49] : Battery Voltage
   // sendBuffer[50] : Battery Voltage
   // sendBuffer[51] : Paused
   // sendBuffer[52] : Last order 1
   // sendBuffer[53] : Last order 2
   // sendBuffer[54] : Current order 1
   // sendBuffer[55] : Current order 2
   // sendBuffer[56] : Last finished 1
   // sendBuffer[57] : Last Finished 2
   // sendBuffer[58] : CS
   // sendBuffer[59] : ETX
   // receiveBuffer[0] : STX
   // receiveBuffer[1] : Size (length of payload)
   // receiveBuffer[2] : Type
   // receiveBuffer[3] : Request ID 1
   // receiveBuffer[4] : Request ID 2
END_DATA_BLOCK

DATA_BLOCK "TCP_IP_Shuttle_DB_13"   // DB387
{ S7_Optimized_Access := 'TRUE' }
VERSION : 0.1
// stored: AutoNumber true, DBAccessibleFromOPCUA true, IsOnlyStoredInLoadMemory false, IsRetainMemResEnabled false, IsWriteProtectedInAS false, MemoryReserve 100
   VAR
      enable : Bool := TRUE;
      send : Bool;
      sendDataLength : UDInt := 0;
      receiveDataLength : UDInt := 16#FFFF_FFFF;
   END_VAR
   VAR RETAIN
      tcpConfig : "LCom_typeConfig";
   END_VAR
   VAR
      tcpDiagnostics { S7_SetPoint := 'True'} : "LCom_typeDiagnostics";
      sendBuffer { S7_SetPoint := 'True'} : Array[0..59] of Byte;
      SendBufferSize : UInt := 60;
      receiveBuffer : Array[0..27] of Byte;
      receiveBufferSize : UInt := 28;
      connected : Bool;
      sending : Bool;
      dataReceived : Bool;
      receivedDataLength : UDInt;
      busy : Bool;
      error : Bool;
      status : Word;
   END_VAR
BEGIN
   tcpConfig.connection.interfaceID := 65164;
   tcpConfig.connection.connectionID := 113;
   tcpConfig.connection.comService := 1;
   tcpConfig.connection.isClient := False;
   tcpConfig.connection.connectType := 1;
   tcpConfig.connection.localPort := 4013;
   tcpConfig.connection.partnerPort := 4013;
   tcpConfig.connection.partnerIP.ADDR[1] := 10;
   tcpConfig.connection.partnerIP.ADDR[2] := 0;
   tcpConfig.connection.partnerIP.ADDR[3] := 34;
   tcpConfig.connection.partnerIP.ADDR[4] := 223;
   tcpConfig.connection.acceptUnknownPartner := TRUE;
   tcpConfig.connection.lifeSignCycleTime := T#1s;
   // sendBuffer[0] : STX
   // sendBuffer[1] : Size
   // sendBuffer[2] : Type
   // sendBuffer[3] : Request ID 1
   // sendBuffer[4] : Request ID 2
   // sendBuffer[5] : PID 1
   // sendBuffer[6] : PID 2
   // sendBuffer[7] : PID 3
   // sendBuffer[8] : PID 4
   // sendBuffer[9] : DID 1
   // sendBuffer[10] : DID 2
   // sendBuffer[11] : DID 3
   // sendBuffer[12] : DID 4
   // sendBuffer[13] : Distance remaining 1
   // sendBuffer[14] : Distance remaining 2
   // sendBuffer[15] : X
   // sendBuffer[16] : X
   // sendBuffer[17] : X
   // sendBuffer[18] : X
   // sendBuffer[19] : Y
   // sendBuffer[20] : Y
   // sendBuffer[21] : Y
   // sendBuffer[22] : Y
   // sendBuffer[23] : Floor
   // sendBuffer[24] : Mode
   // sendBuffer[25] : State
   // sendBuffer[26] : Load State
   // sendBuffer[27] : E1
   // sendBuffer[28] : E1
   // sendBuffer[29] : E2
   // sendBuffer[30] : E2
   // sendBuffer[31] : E3
   // sendBuffer[32] : E3
   // sendBuffer[33] : E4
   // sendBuffer[34] : E4
   // sendBuffer[35] : E5
   // sendBuffer[36] : E5
   // sendBuffer[37] : E6
   // sendBuffer[38] : E6
   // sendBuffer[39] : I1
   // sendBuffer[40] : I1
   // sendBuffer[41] : Q1
   // sendBuffer[42] : Q1
   // sendBuffer[43] : Barcode 1
   // sendBuffer[44] : Barcode 2
   // sendBuffer[45] : Barcode 3
   // sendBuffer[46] : Barcode 4
   // sendBuffer[47] : Pallet Type
   // sendBuffer[48] : Energy Level
   // sendBuffer[49] : Battery Voltage
   // sendBuffer[50] : Battery Voltage
   // sendBuffer[51] : Paused
   // sendBuffer[52] : Last order 1
   // sendBuffer[53] : Last order 2
   // sendBuffer[54] : Current order 1
   // sendBuffer[55] : Current order 2
   // sendBuffer[56] : Last finished 1
   // sendBuffer[57] : Last Finished 2
   // sendBuffer[58] : CS
   // sendBuffer[59] : ETX
   // receiveBuffer[0] : STX
   // receiveBuffer[1] : Size (length of payload)
   // receiveBuffer[2] : Type
   // receiveBuffer[3] : Request ID 1
   // receiveBuffer[4] : Request ID 2
END_DATA_BLOCK

DATA_BLOCK "TCP_IP_Shuttle_DB_14"   // DB378
{ S7_Optimized_Access := 'TRUE' }
VERSION : 0.1
// stored: AutoNumber true, DBAccessibleFromOPCUA true, IsOnlyStoredInLoadMemory false, IsRetainMemResEnabled false, IsWriteProtectedInAS false, MemoryReserve 100
   VAR
      enable : Bool := TRUE;
      send : Bool;
      sendDataLength : UDInt := 0;
      receiveDataLength : UDInt := 16#FFFF_FFFF;
   END_VAR
   VAR RETAIN
      tcpConfig : "LCom_typeConfig";
   END_VAR
   VAR
      tcpDiagnostics { S7_SetPoint := 'True'} : "LCom_typeDiagnostics";
      sendBuffer { S7_SetPoint := 'True'} : Array[0..59] of Byte;
      SendBufferSize : UInt := 60;
      receiveBuffer : Array[0..27] of Byte;
      receiveBufferSize : UInt := 28;
      connected : Bool;
      sending : Bool;
      dataReceived : Bool;
      receivedDataLength : UDInt;
      busy : Bool;
      error : Bool;
      status : Word;
   END_VAR
BEGIN
   tcpConfig.connection.interfaceID := 65164;
   tcpConfig.connection.connectionID := 114;
   tcpConfig.connection.comService := 1;
   tcpConfig.connection.isClient := False;
   tcpConfig.connection.connectType := 1;
   tcpConfig.connection.localPort := 4014;
   tcpConfig.connection.partnerPort := 4014;
   tcpConfig.connection.partnerIP.ADDR[1] := 10;
   tcpConfig.connection.partnerIP.ADDR[2] := 0;
   tcpConfig.connection.partnerIP.ADDR[3] := 34;
   tcpConfig.connection.partnerIP.ADDR[4] := 224;
   tcpConfig.connection.acceptUnknownPartner := TRUE;
   tcpConfig.connection.lifeSignCycleTime := T#1s;
   // sendBuffer[0] : STX
   // sendBuffer[1] : Size
   // sendBuffer[2] : Type
   // sendBuffer[3] : Request ID 1
   // sendBuffer[4] : Request ID 2
   // sendBuffer[5] : PID 1
   // sendBuffer[6] : PID 2
   // sendBuffer[7] : PID 3
   // sendBuffer[8] : PID 4
   // sendBuffer[9] : DID 1
   // sendBuffer[10] : DID 2
   // sendBuffer[11] : DID 3
   // sendBuffer[12] : DID 4
   // sendBuffer[13] : Distance remaining 1
   // sendBuffer[14] : Distance remaining 2
   // sendBuffer[15] : X
   // sendBuffer[16] : X
   // sendBuffer[17] : X
   // sendBuffer[18] : X
   // sendBuffer[19] : Y
   // sendBuffer[20] : Y
   // sendBuffer[21] : Y
   // sendBuffer[22] : Y
   // sendBuffer[23] : Floor
   // sendBuffer[24] : Mode
   // sendBuffer[25] : State
   // sendBuffer[26] : Load State
   // sendBuffer[27] : E1
   // sendBuffer[28] : E1
   // sendBuffer[29] : E2
   // sendBuffer[30] : E2
   // sendBuffer[31] : E3
   // sendBuffer[32] : E3
   // sendBuffer[33] : E4
   // sendBuffer[34] : E4
   // sendBuffer[35] : E5
   // sendBuffer[36] : E5
   // sendBuffer[37] : E6
   // sendBuffer[38] : E6
   // sendBuffer[39] : I1
   // sendBuffer[40] : I1
   // sendBuffer[41] : Q1
   // sendBuffer[42] : Q1
   // sendBuffer[43] : Barcode 1
   // sendBuffer[44] : Barcode 2
   // sendBuffer[45] : Barcode 3
   // sendBuffer[46] : Barcode 4
   // sendBuffer[47] : Pallet Type
   // sendBuffer[48] : Energy Level
   // sendBuffer[49] : Battery Voltage
   // sendBuffer[50] : Battery Voltage
   // sendBuffer[51] : Paused
   // sendBuffer[52] : Last order 1
   // sendBuffer[53] : Last order 2
   // sendBuffer[54] : Current order 1
   // sendBuffer[55] : Current order 2
   // sendBuffer[56] : Last finished 1
   // sendBuffer[57] : Last Finished 2
   // sendBuffer[58] : CS
   // sendBuffer[59] : ETX
   // receiveBuffer[0] : STX
   // receiveBuffer[1] : Size (length of payload)
   // receiveBuffer[2] : Type
   // receiveBuffer[3] : Request ID 1
   // receiveBuffer[4] : Request ID 2
END_DATA_BLOCK

DATA_BLOCK "TCP_IP_Shuttle_DB_15"   // DB389
{ S7_Optimized_Access := 'TRUE' }
VERSION : 0.1
// stored: AutoNumber true, DBAccessibleFromOPCUA true, IsOnlyStoredInLoadMemory false, IsRetainMemResEnabled false, IsWriteProtectedInAS false, MemoryReserve 100
   VAR
      enable : Bool := TRUE;
      send : Bool;
      sendDataLength : UDInt := 0;
      receiveDataLength : UDInt := 16#FFFF_FFFF;
   END_VAR
   VAR RETAIN
      tcpConfig : "LCom_typeConfig";
   END_VAR
   VAR
      tcpDiagnostics { S7_SetPoint := 'True'} : "LCom_typeDiagnostics";
      sendBuffer { S7_SetPoint := 'True'} : Array[0..59] of Byte;
      SendBufferSize : UInt := 60;
      receiveBuffer : Array[0..27] of Byte;
      receiveBufferSize : UInt := 28;
      connected : Bool;
      sending : Bool;
      dataReceived : Bool;
      receivedDataLength : UDInt;
      busy : Bool;
      error : Bool;
      status : Word;
   END_VAR
BEGIN
   tcpConfig.connection.interfaceID := 65164;
   tcpConfig.connection.connectionID := 115;
   tcpConfig.connection.comService := 1;
   tcpConfig.connection.isClient := False;
   tcpConfig.connection.connectType := 1;
   tcpConfig.connection.localPort := 4015;
   tcpConfig.connection.partnerPort := 4015;
   tcpConfig.connection.partnerIP.ADDR[1] := 10;
   tcpConfig.connection.partnerIP.ADDR[2] := 0;
   tcpConfig.connection.partnerIP.ADDR[3] := 34;
   tcpConfig.connection.partnerIP.ADDR[4] := 225;
   tcpConfig.connection.acceptUnknownPartner := TRUE;
   tcpConfig.connection.lifeSignCycleTime := T#1s;
   // sendBuffer[0] : STX
   // sendBuffer[1] : Size
   // sendBuffer[2] : Type
   // sendBuffer[3] : Request ID 1
   // sendBuffer[4] : Request ID 2
   // sendBuffer[5] : PID 1
   // sendBuffer[6] : PID 2
   // sendBuffer[7] : PID 3
   // sendBuffer[8] : PID 4
   // sendBuffer[9] : DID 1
   // sendBuffer[10] : DID 2
   // sendBuffer[11] : DID 3
   // sendBuffer[12] : DID 4
   // sendBuffer[13] : Distance remaining 1
   // sendBuffer[14] : Distance remaining 2
   // sendBuffer[15] : X
   // sendBuffer[16] : X
   // sendBuffer[17] : X
   // sendBuffer[18] : X
   // sendBuffer[19] : Y
   // sendBuffer[20] : Y
   // sendBuffer[21] : Y
   // sendBuffer[22] : Y
   // sendBuffer[23] : Floor
   // sendBuffer[24] : Mode
   // sendBuffer[25] : State
   // sendBuffer[26] : Load State
   // sendBuffer[27] : E1
   // sendBuffer[28] : E1
   // sendBuffer[29] : E2
   // sendBuffer[30] : E2
   // sendBuffer[31] : E3
   // sendBuffer[32] : E3
   // sendBuffer[33] : E4
   // sendBuffer[34] : E4
   // sendBuffer[35] : E5
   // sendBuffer[36] : E5
   // sendBuffer[37] : E6
   // sendBuffer[38] : E6
   // sendBuffer[39] : I1
   // sendBuffer[40] : I1
   // sendBuffer[41] : Q1
   // sendBuffer[42] : Q1
   // sendBuffer[43] : Barcode 1
   // sendBuffer[44] : Barcode 2
   // sendBuffer[45] : Barcode 3
   // sendBuffer[46] : Barcode 4
   // sendBuffer[47] : Pallet Type
   // sendBuffer[48] : Energy Level
   // sendBuffer[49] : Battery Voltage
   // sendBuffer[50] : Battery Voltage
   // sendBuffer[51] : Paused
   // sendBuffer[52] : Last order 1
   // sendBuffer[53] : Last order 2
   // sendBuffer[54] : Current order 1
   // sendBuffer[55] : Current order 2
   // sendBuffer[56] : Last finished 1
   // sendBuffer[57] : Last Finished 2
   // sendBuffer[58] : CS
   // sendBuffer[59] : ETX
   // receiveBuffer[0] : STX
   // receiveBuffer[1] : Size (length of payload)
   // receiveBuffer[2] : Type
   // receiveBuffer[3] : Request ID 1
   // receiveBuffer[4] : Request ID 2
END_DATA_BLOCK

DATA_BLOCK "TCP_IP_Shuttle_DB_16"   // DB381
{ S7_Optimized_Access := 'TRUE' }
VERSION : 0.1
// stored: AutoNumber true, DBAccessibleFromOPCUA true, IsOnlyStoredInLoadMemory false, IsRetainMemResEnabled false, IsWriteProtectedInAS false, MemoryReserve 100
   VAR
      enable : Bool := TRUE;
      send : Bool;
      sendDataLength : UDInt := 0;
      receiveDataLength : UDInt := 16#FFFF_FFFF;
   END_VAR
   VAR RETAIN
      tcpConfig : "LCom_typeConfig";
   END_VAR
   VAR
      tcpDiagnostics { S7_SetPoint := 'True'} : "LCom_typeDiagnostics";
      sendBuffer { S7_SetPoint := 'True'} : Array[0..59] of Byte;
      SendBufferSize : UInt := 60;
      receiveBuffer : Array[0..27] of Byte;
      receiveBufferSize : UInt := 28;
      connected : Bool;
      sending : Bool;
      dataReceived : Bool;
      receivedDataLength : UDInt;
      busy : Bool;
      error : Bool;
      status : Word;
   END_VAR
BEGIN
   tcpConfig.connection.interfaceID := 65164;
   tcpConfig.connection.connectionID := 116;
   tcpConfig.connection.comService := 1;
   tcpConfig.connection.isClient := False;
   tcpConfig.connection.connectType := 1;
   tcpConfig.connection.localPort := 4016;
   tcpConfig.connection.partnerPort := 4016;
   tcpConfig.connection.partnerIP.ADDR[1] := 10;
   tcpConfig.connection.partnerIP.ADDR[2] := 0;
   tcpConfig.connection.partnerIP.ADDR[3] := 34;
   tcpConfig.connection.partnerIP.ADDR[4] := 226;
   tcpConfig.connection.acceptUnknownPartner := TRUE;
   tcpConfig.connection.lifeSignCycleTime := T#1s;
   // sendBuffer[0] : STX
   // sendBuffer[1] : Size
   // sendBuffer[2] : Type
   // sendBuffer[3] : Request ID 1
   // sendBuffer[4] : Request ID 2
   // sendBuffer[5] : PID 1
   // sendBuffer[6] : PID 2
   // sendBuffer[7] : PID 3
   // sendBuffer[8] : PID 4
   // sendBuffer[9] : DID 1
   // sendBuffer[10] : DID 2
   // sendBuffer[11] : DID 3
   // sendBuffer[12] : DID 4
   // sendBuffer[13] : Distance remaining 1
   // sendBuffer[14] : Distance remaining 2
   // sendBuffer[15] : X
   // sendBuffer[16] : X
   // sendBuffer[17] : X
   // sendBuffer[18] : X
   // sendBuffer[19] : Y
   // sendBuffer[20] : Y
   // sendBuffer[21] : Y
   // sendBuffer[22] : Y
   // sendBuffer[23] : Floor
   // sendBuffer[24] : Mode
   // sendBuffer[25] : State
   // sendBuffer[26] : Load State
   // sendBuffer[27] : E1
   // sendBuffer[28] : E1
   // sendBuffer[29] : E2
   // sendBuffer[30] : E2
   // sendBuffer[31] : E3
   // sendBuffer[32] : E3
   // sendBuffer[33] : E4
   // sendBuffer[34] : E4
   // sendBuffer[35] : E5
   // sendBuffer[36] : E5
   // sendBuffer[37] : E6
   // sendBuffer[38] : E6
   // sendBuffer[39] : I1
   // sendBuffer[40] : I1
   // sendBuffer[41] : Q1
   // sendBuffer[42] : Q1
   // sendBuffer[43] : Barcode 1
   // sendBuffer[44] : Barcode 2
   // sendBuffer[45] : Barcode 3
   // sendBuffer[46] : Barcode 4
   // sendBuffer[47] : Pallet Type
   // sendBuffer[48] : Energy Level
   // sendBuffer[49] : Battery Voltage
   // sendBuffer[50] : Battery Voltage
   // sendBuffer[51] : Paused
   // sendBuffer[52] : Last order 1
   // sendBuffer[53] : Last order 2
   // sendBuffer[54] : Current order 1
   // sendBuffer[55] : Current order 2
   // sendBuffer[56] : Last finished 1
   // sendBuffer[57] : Last Finished 2
   // sendBuffer[58] : CS
   // sendBuffer[59] : ETX
   // receiveBuffer[0] : STX
   // receiveBuffer[1] : Size (length of payload)
   // receiveBuffer[2] : Type
   // receiveBuffer[3] : Request ID 1
   // receiveBuffer[4] : Request ID 2
END_DATA_BLOCK

DATA_BLOCK "TCP_IP_Shuttle_DB_17"   // DB379
{ S7_Optimized_Access := 'TRUE' }
VERSION : 0.1
// stored: AutoNumber true, DBAccessibleFromOPCUA true, IsOnlyStoredInLoadMemory false, IsRetainMemResEnabled false, IsWriteProtectedInAS false, MemoryReserve 100
   VAR
      enable : Bool := TRUE;
      send : Bool;
      sendDataLength : UDInt := 0;
      receiveDataLength : UDInt := 16#FFFF_FFFF;
   END_VAR
   VAR RETAIN
      tcpConfig : "LCom_typeConfig";
   END_VAR
   VAR
      tcpDiagnostics { S7_SetPoint := 'True'} : "LCom_typeDiagnostics";
      sendBuffer { S7_SetPoint := 'True'} : Array[0..59] of Byte;
      SendBufferSize : UInt := 60;
      receiveBuffer : Array[0..27] of Byte;
      receiveBufferSize : UInt := 28;
      connected : Bool;
      sending : Bool;
      dataReceived : Bool;
      receivedDataLength : UDInt;
      busy : Bool;
      error : Bool;
      status : Word;
   END_VAR
BEGIN
   tcpConfig.connection.interfaceID := 65164;
   tcpConfig.connection.connectionID := 117;
   tcpConfig.connection.comService := 1;
   tcpConfig.connection.isClient := False;
   tcpConfig.connection.connectType := 1;
   tcpConfig.connection.localPort := 4017;
   tcpConfig.connection.partnerPort := 4017;
   tcpConfig.connection.partnerIP.ADDR[1] := 10;
   tcpConfig.connection.partnerIP.ADDR[2] := 0;
   tcpConfig.connection.partnerIP.ADDR[3] := 34;
   tcpConfig.connection.partnerIP.ADDR[4] := 227;
   tcpConfig.connection.acceptUnknownPartner := TRUE;
   tcpConfig.connection.lifeSignCycleTime := T#1s;
   // sendBuffer[0] : STX
   // sendBuffer[1] : Size
   // sendBuffer[2] : Type
   // sendBuffer[3] : Request ID 1
   // sendBuffer[4] : Request ID 2
   // sendBuffer[5] : PID 1
   // sendBuffer[6] : PID 2
   // sendBuffer[7] : PID 3
   // sendBuffer[8] : PID 4
   // sendBuffer[9] : DID 1
   // sendBuffer[10] : DID 2
   // sendBuffer[11] : DID 3
   // sendBuffer[12] : DID 4
   // sendBuffer[13] : Distance remaining 1
   // sendBuffer[14] : Distance remaining 2
   // sendBuffer[15] : X
   // sendBuffer[16] : X
   // sendBuffer[17] : X
   // sendBuffer[18] : X
   // sendBuffer[19] : Y
   // sendBuffer[20] : Y
   // sendBuffer[21] : Y
   // sendBuffer[22] : Y
   // sendBuffer[23] : Floor
   // sendBuffer[24] : Mode
   // sendBuffer[25] : State
   // sendBuffer[26] : Load State
   // sendBuffer[27] : E1
   // sendBuffer[28] : E1
   // sendBuffer[29] : E2
   // sendBuffer[30] : E2
   // sendBuffer[31] : E3
   // sendBuffer[32] : E3
   // sendBuffer[33] : E4
   // sendBuffer[34] : E4
   // sendBuffer[35] : E5
   // sendBuffer[36] : E5
   // sendBuffer[37] : E6
   // sendBuffer[38] : E6
   // sendBuffer[39] : I1
   // sendBuffer[40] : I1
   // sendBuffer[41] : Q1
   // sendBuffer[42] : Q1
   // sendBuffer[43] : Barcode 1
   // sendBuffer[44] : Barcode 2
   // sendBuffer[45] : Barcode 3
   // sendBuffer[46] : Barcode 4
   // sendBuffer[47] : Pallet Type
   // sendBuffer[48] : Energy Level
   // sendBuffer[49] : Battery Voltage
   // sendBuffer[50] : Battery Voltage
   // sendBuffer[51] : Paused
   // sendBuffer[52] : Last order 1
   // sendBuffer[53] : Last order 2
   // sendBuffer[54] : Current order 1
   // sendBuffer[55] : Current order 2
   // sendBuffer[56] : Last finished 1
   // sendBuffer[57] : Last Finished 2
   // sendBuffer[58] : CS
   // sendBuffer[59] : ETX
   // receiveBuffer[0] : STX
   // receiveBuffer[1] : Size (length of payload)
   // receiveBuffer[2] : Type
   // receiveBuffer[3] : Request ID 1
   // receiveBuffer[4] : Request ID 2
END_DATA_BLOCK

DATA_BLOCK "TCP_IP_Shuttle_DB_18"   // DB240
{ S7_Optimized_Access := 'TRUE' }
VERSION : 0.1
// stored: AutoNumber true, DBAccessibleFromOPCUA true, IsOnlyStoredInLoadMemory false, IsRetainMemResEnabled false, IsWriteProtectedInAS false, MemoryReserve 100
   VAR
      enable : Bool := TRUE;
      send : Bool;
      sendDataLength : UDInt := 0;
      receiveDataLength : UDInt := 16#FFFF_FFFF;
   END_VAR
   VAR RETAIN
      tcpConfig : "LCom_typeConfig";
   END_VAR
   VAR
      tcpDiagnostics { S7_SetPoint := 'True'} : "LCom_typeDiagnostics";
      sendBuffer { S7_SetPoint := 'True'} : Array[0..59] of Byte;
      SendBufferSize : UInt := 60;
      receiveBuffer : Array[0..27] of Byte;
      receiveBufferSize : UInt := 28;
      connected : Bool;
      sending : Bool;
      dataReceived : Bool;
      receivedDataLength : UDInt;
      busy : Bool;
      error : Bool;
      status : Word;
   END_VAR
BEGIN
   tcpConfig.connection.interfaceID := 65164;
   tcpConfig.connection.connectionID := 118;
   tcpConfig.connection.comService := 1;
   tcpConfig.connection.isClient := False;
   tcpConfig.connection.connectType := 1;
   tcpConfig.connection.localPort := 4018;
   tcpConfig.connection.partnerPort := 4018;
   tcpConfig.connection.partnerIP.ADDR[1] := 10;
   tcpConfig.connection.partnerIP.ADDR[2] := 0;
   tcpConfig.connection.partnerIP.ADDR[3] := 34;
   tcpConfig.connection.partnerIP.ADDR[4] := 228;
   tcpConfig.connection.acceptUnknownPartner := TRUE;
   tcpConfig.connection.lifeSignCycleTime := T#1s;
   // sendBuffer[0] : STX
   // sendBuffer[1] : Size
   // sendBuffer[2] : Type
   // sendBuffer[3] : Request ID 1
   // sendBuffer[4] : Request ID 2
   // sendBuffer[5] : PID 1
   // sendBuffer[6] : PID 2
   // sendBuffer[7] : PID 3
   // sendBuffer[8] : PID 4
   // sendBuffer[9] : DID 1
   // sendBuffer[10] : DID 2
   // sendBuffer[11] : DID 3
   // sendBuffer[12] : DID 4
   // sendBuffer[13] : Distance remaining 1
   // sendBuffer[14] : Distance remaining 2
   // sendBuffer[15] : X
   // sendBuffer[16] : X
   // sendBuffer[17] : X
   // sendBuffer[18] : X
   // sendBuffer[19] : Y
   // sendBuffer[20] : Y
   // sendBuffer[21] : Y
   // sendBuffer[22] : Y
   // sendBuffer[23] : Floor
   // sendBuffer[24] : Mode
   // sendBuffer[25] : State
   // sendBuffer[26] : Load State
   // sendBuffer[27] : E1
   // sendBuffer[28] : E1
   // sendBuffer[29] : E2
   // sendBuffer[30] : E2
   // sendBuffer[31] : E3
   // sendBuffer[32] : E3
   // sendBuffer[33] : E4
   // sendBuffer[34] : E4
   // sendBuffer[35] : E5
   // sendBuffer[36] : E5
   // sendBuffer[37] : E6
   // sendBuffer[38] : E6
   // sendBuffer[39] : I1
   // sendBuffer[40] : I1
   // sendBuffer[41] : Q1
   // sendBuffer[42] : Q1
   // sendBuffer[43] : Barcode 1
   // sendBuffer[44] : Barcode 2
   // sendBuffer[45] : Barcode 3
   // sendBuffer[46] : Barcode 4
   // sendBuffer[47] : Pallet Type
   // sendBuffer[48] : Energy Level
   // sendBuffer[49] : Battery Voltage
   // sendBuffer[50] : Battery Voltage
   // sendBuffer[51] : Paused
   // sendBuffer[52] : Last order 1
   // sendBuffer[53] : Last order 2
   // sendBuffer[54] : Current order 1
   // sendBuffer[55] : Current order 2
   // sendBuffer[56] : Last finished 1
   // sendBuffer[57] : Last Finished 2
   // sendBuffer[58] : CS
   // sendBuffer[59] : ETX
   // receiveBuffer[0] : STX
   // receiveBuffer[1] : Size (length of payload)
   // receiveBuffer[2] : Type
   // receiveBuffer[3] : Request ID 1
   // receiveBuffer[4] : Request ID 2
END_DATA_BLOCK

DATA_BLOCK "TCP_IP_Shuttle_DB_19"   // DB239
{ S7_Optimized_Access := 'TRUE' }
VERSION : 0.1
// stored: AutoNumber true, DBAccessibleFromOPCUA true, IsOnlyStoredInLoadMemory false, IsRetainMemResEnabled false, IsWriteProtectedInAS false, MemoryReserve 100
   VAR
      enable : Bool := TRUE;
      send : Bool;
      sendDataLength : UDInt := 0;
      receiveDataLength : UDInt := 16#FFFF_FFFF;
   END_VAR
   VAR RETAIN
      tcpConfig : "LCom_typeConfig";
   END_VAR
   VAR
      tcpDiagnostics { S7_SetPoint := 'True'} : "LCom_typeDiagnostics";
      sendBuffer { S7_SetPoint := 'True'} : Array[0..59] of Byte;
      SendBufferSize : UInt := 60;
      receiveBuffer : Array[0..27] of Byte;
      receiveBufferSize : UInt := 28;
      connected : Bool;
      sending : Bool;
      dataReceived : Bool;
      receivedDataLength : UDInt;
      busy : Bool;
      error : Bool;
      status : Word;
   END_VAR
BEGIN
   tcpConfig.connection.interfaceID := 65164;
   tcpConfig.connection.connectionID := 119;
   tcpConfig.connection.comService := 1;
   tcpConfig.connection.isClient := False;
   tcpConfig.connection.connectType := 1;
   tcpConfig.connection.localPort := 4019;
   tcpConfig.connection.partnerPort := 4019;
   tcpConfig.connection.partnerIP.ADDR[1] := 10;
   tcpConfig.connection.partnerIP.ADDR[2] := 0;
   tcpConfig.connection.partnerIP.ADDR[3] := 34;
   tcpConfig.connection.partnerIP.ADDR[4] := 229;
   tcpConfig.connection.acceptUnknownPartner := TRUE;
   tcpConfig.connection.lifeSignCycleTime := T#1s;
   // sendBuffer[0] : STX
   // sendBuffer[1] : Size
   // sendBuffer[2] : Type
   // sendBuffer[3] : Request ID 1
   // sendBuffer[4] : Request ID 2
   // sendBuffer[5] : PID 1
   // sendBuffer[6] : PID 2
   // sendBuffer[7] : PID 3
   // sendBuffer[8] : PID 4
   // sendBuffer[9] : DID 1
   // sendBuffer[10] : DID 2
   // sendBuffer[11] : DID 3
   // sendBuffer[12] : DID 4
   // sendBuffer[13] : Distance remaining 1
   // sendBuffer[14] : Distance remaining 2
   // sendBuffer[15] : X
   // sendBuffer[16] : X
   // sendBuffer[17] : X
   // sendBuffer[18] : X
   // sendBuffer[19] : Y
   // sendBuffer[20] : Y
   // sendBuffer[21] : Y
   // sendBuffer[22] : Y
   // sendBuffer[23] : Floor
   // sendBuffer[24] : Mode
   // sendBuffer[25] : State
   // sendBuffer[26] : Load State
   // sendBuffer[27] : E1
   // sendBuffer[28] : E1
   // sendBuffer[29] : E2
   // sendBuffer[30] : E2
   // sendBuffer[31] : E3
   // sendBuffer[32] : E3
   // sendBuffer[33] : E4
   // sendBuffer[34] : E4
   // sendBuffer[35] : E5
   // sendBuffer[36] : E5
   // sendBuffer[37] : E6
   // sendBuffer[38] : E6
   // sendBuffer[39] : I1
   // sendBuffer[40] : I1
   // sendBuffer[41] : Q1
   // sendBuffer[42] : Q1
   // sendBuffer[43] : Barcode 1
   // sendBuffer[44] : Barcode 2
   // sendBuffer[45] : Barcode 3
   // sendBuffer[46] : Barcode 4
   // sendBuffer[47] : Pallet Type
   // sendBuffer[48] : Energy Level
   // sendBuffer[49] : Battery Voltage
   // sendBuffer[50] : Battery Voltage
   // sendBuffer[51] : Paused
   // sendBuffer[52] : Last order 1
   // sendBuffer[53] : Last order 2
   // sendBuffer[54] : Current order 1
   // sendBuffer[55] : Current order 2
   // sendBuffer[56] : Last finished 1
   // sendBuffer[57] : Last Finished 2
   // sendBuffer[58] : CS
   // sendBuffer[59] : ETX
   // receiveBuffer[0] : STX
   // receiveBuffer[1] : Size (length of payload)
   // receiveBuffer[2] : Type
   // receiveBuffer[3] : Request ID 1
   // receiveBuffer[4] : Request ID 2
END_DATA_BLOCK

DATA_BLOCK "TCP_IP_Shuttle_DB_2"   // DB305
{ S7_Optimized_Access := 'TRUE' }
VERSION : 0.1
// stored: AutoNumber true, DBAccessibleFromOPCUA true, IsOnlyStoredInLoadMemory false, IsRetainMemResEnabled false, IsWriteProtectedInAS false, MemoryReserve 100
   VAR
      enable : Bool := TRUE;
      send : Bool;
      sendDataLength : UDInt := 0;
      receiveDataLength : UDInt := 16#FFFF_FFFF;
   END_VAR
   VAR RETAIN
      tcpConfig : "LCom_typeConfig";
   END_VAR
   VAR
      tcpDiagnostics { S7_SetPoint := 'True'} : "LCom_typeDiagnostics";
      sendBuffer { S7_SetPoint := 'True'} : Array[0..59] of Byte;
      SendBufferSize : UInt := 60;
      receiveBuffer : Array[0..27] of Byte;
      receiveBufferSize : UInt := 28;
      connected : Bool;
      sending : Bool;
      dataReceived : Bool;
      receivedDataLength : UDInt;
      busy : Bool;
      error : Bool;
      status : Word;
   END_VAR
BEGIN
   tcpConfig.connection.interfaceID := 65164;
   tcpConfig.connection.connectionID := 102;
   tcpConfig.connection.comService := 1;
   tcpConfig.connection.isClient := False;
   tcpConfig.connection.connectType := 1;
   tcpConfig.connection.localPort := 4002;
   tcpConfig.connection.partnerPort := 4002;
   tcpConfig.connection.partnerIP.ADDR[1] := 10;
   tcpConfig.connection.partnerIP.ADDR[2] := 0;
   tcpConfig.connection.partnerIP.ADDR[3] := 35;
   tcpConfig.connection.partnerIP.ADDR[4] := 62;
   tcpConfig.connection.acceptUnknownPartner := TRUE;
   tcpConfig.connection.lifeSignCycleTime := T#1s;
   // sendBuffer[0] : STX
   // sendBuffer[1] : Size
   // sendBuffer[2] : Type
   // sendBuffer[3] : Request ID 1
   // sendBuffer[4] : Request ID 2
   // sendBuffer[5] : PID 1
   // sendBuffer[6] : PID 2
   // sendBuffer[7] : PID 3
   // sendBuffer[8] : PID 4
   // sendBuffer[9] : DID 1
   // sendBuffer[10] : DID 2
   // sendBuffer[11] : DID 3
   // sendBuffer[12] : DID 4
   // sendBuffer[13] : Distance remaining 1
   // sendBuffer[14] : Distance remaining 2
   // sendBuffer[15] : X
   // sendBuffer[16] : X
   // sendBuffer[17] : X
   // sendBuffer[18] : X
   // sendBuffer[19] : Y
   // sendBuffer[20] : Y
   // sendBuffer[21] : Y
   // sendBuffer[22] : Y
   // sendBuffer[23] : Floor
   // sendBuffer[24] : Mode
   // sendBuffer[25] : State
   // sendBuffer[26] : Load State
   // sendBuffer[27] : E1
   // sendBuffer[28] : E1
   // sendBuffer[29] : E2
   // sendBuffer[30] : E2
   // sendBuffer[31] : E3
   // sendBuffer[32] : E3
   // sendBuffer[33] : E4
   // sendBuffer[34] : E4
   // sendBuffer[35] : E5
   // sendBuffer[36] : E5
   // sendBuffer[37] : E6
   // sendBuffer[38] : E6
   // sendBuffer[39] : I1
   // sendBuffer[40] : I1
   // sendBuffer[41] : Q1
   // sendBuffer[42] : Q1
   // sendBuffer[43] : Barcode 1
   // sendBuffer[44] : Barcode 2
   // sendBuffer[45] : Barcode 3
   // sendBuffer[46] : Barcode 4
   // sendBuffer[47] : Pallet Type
   // sendBuffer[48] : Energy Level
   // sendBuffer[49] : Battery Voltage
   // sendBuffer[50] : Battery Voltage
   // sendBuffer[51] : Paused
   // sendBuffer[52] : Last order 1
   // sendBuffer[53] : Last order 2
   // sendBuffer[54] : Current order 1
   // sendBuffer[55] : Current order 2
   // sendBuffer[56] : Last finished 1
   // sendBuffer[57] : Last Finished 2
   // sendBuffer[58] : CS
   // sendBuffer[59] : ETX
   // receiveBuffer[0] : STX
   // receiveBuffer[1] : Size (length of payload)
   // receiveBuffer[2] : Type
   // receiveBuffer[3] : Request ID 1
   // receiveBuffer[4] : Request ID 2
END_DATA_BLOCK

